Universal Robots PolyScope program: AdientTorsF_Eol1R.urp

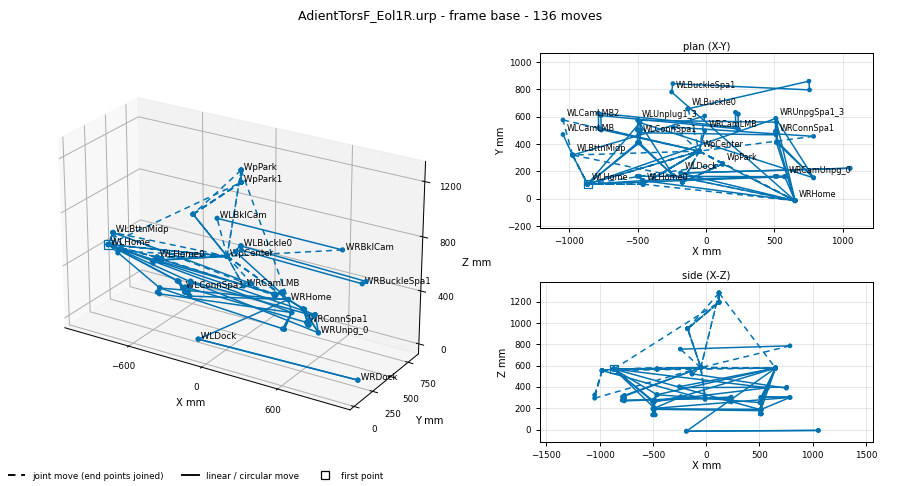
[picture p0: tool path of AdientTorsF_Eol1R.urp in frame base, 136 of 176 moves have a stored position in this frame; points joined in program order, loops and branches not executed]
Program AdientTorsF_Eol1R (installation=EOL_1R directory=/programs createdIn=3.5.1 lastSavedIn=5.26.0 robotSerialNumber=20265101874)
Calibrated DH parameters: a=[0.000042, -0.610949, -0.549442, -0.000024, -0.000005, 0]; d=[0.18065, -32.695743, 7.316343, 25.554022, 0.119806, 0.115349]; alpha=[1.570492, -0.001088, 0.006138, 1.570534, -1.57033, 0]; deltaTheta=[0, 0.058138, -0.334397, 0.276266, -0.000002, 0]
InitVariablesNode variables(variable(name=Abort, expression=False), variable(name=AdapterReady_L, expression=False), variable(name=AdapterReady_R, expression=False), variable(name=CMD_Heartbt_i1, expression=0), variable(name=CMD_Heartbt_i2, expression=0), variable(name=CMD_Program_i1, expression=0), variable(name=CMD_Program_i2, expression=0), variable(name=CMD_Reserve_i1, expression=0), variable(name=CMD_Reserve_i2, expression=0), variable(name=CMD_Timeout_i1, expression=0), variable(name=CMD_Timeout_i2, expression=0), variable(name=CamCorrectnOK, expression=0), variable(name=DEBUG, expression=False), variable(name=D_rel, expression=p[0,0,0,0,0,0]), variable(name=EvtBeep, expression=False), variable(name=EvtDock, expression=0), variable(name=Mute, expression=False), variable(name=P_ini, expression=get_actual_tcp_pose()), variable(name=Parking, expression=0), variable(name=ProgExe, expression=0), variable(name=STS_Heartbeat, expression=False), variable(name=STS_Progress, expression=0), variable(name=STS_Reservation, expression=0), variable(name=SetCameraProg, expression=0))
BeforeStart
  SuppressedNode
    DEBUG := True
  'SW version, to be used to track changes and keep sync of all stations'
  SW_Ver := 1.0
  Folder Scripts [hidden by the author, left out]
  Folder Avoid guidance screen [hidden by the author, left out]
  Call GripperOpen
  GoToHome := True
  Script: socket_open("127.0.0.1",30001)
Robot Program (runOnlyOnce=false)
  Folder Execute Program
    Folder Init
      Wait Condition expression=EvtDock≤0
      Folder Verify adapter ready
        If Di_Docked_L or AI_Gripper<(ivGripSensOpen+0.3)
          AdapterReady_L := False
        If Di_Docked_R or AI_Gripper<(ivGripSensOpen+0.3)
          AdapterReady_R := False
      Folder Go to home pos automatically
        If GoToHome and  not (AdapterReady_L or AdapterReady_R)
          Wait Sleep waitTime=1
          If InRange(P_Flange[0],-1,-0.2) and InRange(P_Flange[1],-0.5,0.5) and InRange(P_Flange[2],0.3,1)
            If AdapterDocked or DEBUG or (AI_Gripper<(ivGripSensOpen+0.3))
              MoveJ speed 120 deg/s, acceleration 500 deg/s^2 (useActiveTCP=false positionType=JointAngles optimoveEnabled=false optiMoveSpeed=0.3 optiMoveAcceleration=0.09) tcp=t0_Flange; feature=Base
                Waypoint WLHome: TCP in base x=-866.235 y=106.553 z=568.537 mm, rx=3.1416 ry=0 rz=0 rad; joints [-18.569, -73.864, 82.281, -98.358, -89.699, -108.526] deg; TCP offset x=0 y=0 z=0 mm, rx=0 ry=0 rz=3.1416 rad
            Else 
              Popup Error (haltProgram=false message=Adapter must be docked inputType=Text)
              Halt
          ElseIf AtCenterPos
            MoveJ speed 120 deg/s, acceleration 500 deg/s^2 (useActiveTCP=true positionType=JointAngles optimoveEnabled=false optiMoveSpeed=0.3 optiMoveAcceleration=0.09) feature=Base
              Waypoint WpCenter: TCP in base x=-50 y=348.529 z=581.932 mm, rx=0 ry=3.1416 rz=0 rad; joints [-111.545, -128.858, 124.717, -85.8, -89.657, -21.591] deg; TCP offset x=0 y=0 z=0 mm, rx=0 ry=0 rz=3.1416 rad
          ElseIf AtParkPos
            MoveJ speed 120 deg/s, acceleration 500 deg/s^2 (useActiveTCP=true positionType=JointAngles optimoveEnabled=false optiMoveSpeed=0.3 optiMoveAcceleration=0.09) feature=Base
              Waypoint WpPark: TCP in base x=121.203 y=255.21 z=1282.913 mm, rx=-1.7636 ry=-1.7554 rz=-0.7332 rad; joints [-180, -89.998, -0.001, 0.001, -45, 0] deg; TCP offset x=0 y=0 z=0 mm, rx=0 ry=0 rz=3.1416 rad
          ElseIf InRange(P_Flange[0],0.2,1.2) and InRange(P_Flange[1],-0.5,0.5) and InRange(P_Flange[2],0.3,1)
            If AdapterDocked or DEBUG or (AI_Gripper<(ivGripSensOpen+0.3))
              MoveJ speed 120 deg/s, acceleration 500 deg/s^2 (useActiveTCP=true positionType=JointAngles optimoveEnabled=false optiMoveSpeed=0.3 optiMoveAcceleration=0.09) feature=Base
                Waypoint WRHome: TCP in base x=651.404 y=-14.037 z=577.942 mm, rx=3.1416 ry=0 rz=0 rad; joints [-196.798, -95.185, 104.834, -99.59, -89.673, 73.253] deg
            Else 
              Popup Error (haltProgram=false message=Adapter must be docked inputType=Text)
              Halt
          Else 
            Popup Error (haltProgram=false message=Illegal position. Adjust arm to open space in front of the backrest, or [Move]->[Home] inputType=Text)
            Halt
        GoToHome := False
      If DEBUG
        'Popup window with program selection'
        ProgExe :=  (valueSource=Operator message=Program number? valueType=Integer)
      If ProgExe>0
        Folder Init
          Mute := False
          Wait Condition expression=not GoToHome
          If In(ProgExe,[11,12,14])
            AdapterReady_R := False
          ElseIf In(ProgExe,[51,52,54])
            AdapterReady_L := False
          Else 
            AdapterReady_L := False
            AdapterReady_R := False
    Folder Programs
      If InRange(ProgExe,1,99)
        Folder Undock
          If In(ProgExe,[11,51])
            Script: Report(1)
            Folder AtHome?
              Timer (action=Reset) variable(name=T_Timeout)
              Timer (action=Start) variable=T_Timeout
              Wait Condition expression=AtHomePos or T_Timeout>5
              If not AtHomePos
                Script: Report(90)
            If Progress_run() and  not AdapterDocked
              Script: Report(94)
            If Progress_run()
              Folder Undock
                MoveL speed 1000 mm/s, acceleration 3000 mm/s^2 (useActiveTCP=false optimoveEnabled=false optiMoveSpeed=0.3 optiMoveAcceleration=0.09) tcp=t2_Gripper; feature=Base
                  Call GripperOpenQuick
                  If False
                    Waypoint WLDock: TCP in base x=-185.159 y=188.226 z=-15.087 mm, rx=1.8903 ry=-1.8549 rz=-0.6082 rad; joints [-63.281, -90.699, 161.642, -179.168, -58.985, -58.884] deg; TCP offset x=0 y=260 z=74 mm, rx=0 ry=0 rz=3.1416 rad
                    Waypoint WRDock: TCP in base x=1053.302 y=223.512 z=-7.7 mm, rx=1.9028 ry=-1.8549 rz=-0.594 rad; joints [-177.46, -52.491, 84.331, -87.181, -88.23, 180.6] deg
                  If ProgExe<50
                    WpDock := WLDock
                    WpHome := WLHome
                  Else 
                    WpDock := WRDock
                    WpHome := WRHome
                  Wp := pose_trans(WpDock, p[0,0.175,-0.1,0,0,0])
                  Waypoint Variable (Variable): motionParameters(blendRadius=0.05); variable=Wp
                  Call GripperOpen
                  Wp := pose_trans(WpDock, p[0,0.075,0.01,0,0,0])
                  Waypoint Variable (Variable): motionParameters(blendRadius=0.01); variable=Wp
                  Wp := pose_trans(WpDock, p[0,0.055,0,0,0,0])
                  Waypoint Variable (Variable): motionParameters(blendRadius=0.01); variable=Wp
                  Waypoint Variable (Variable): variable=WpDock
                  Call GripperClose
                  Wp := pose_trans(WpDock, p[0,0.25,0,0,0,0])
                  Waypoint Variable (Variable): variable=Wp
                If ProgExe<50
                  AdapterReady_L := True
                Else 
                  AdapterReady_R := True
                Script: Report(50)
            Script: Report(50)
        Folder Connect
          If In(ProgExe,[12,14,52,54])
            Script: Report(1)
            If ProgExe<50 and AdapterReady_L
              Undock := False
            ElseIf ProgExe≥50 and AdapterReady_R
              Undock := False
            Else 
              Undock := True
              Folder AtHome? [hidden by the author, left out]
              If Progress_run() and  not AdapterDocked
                Script: Report(94)
            If Progress_run()
              Folder Undock
                If Undock
                  MoveL speed 1000 mm/s, acceleration 3000 mm/s^2 (useActiveTCP=false optimoveEnabled=false optiMoveSpeed=0.3 optiMoveAcceleration=0.09) tcp=t2_Gripper; feature=Base
                    Call GripperOpenQuick
                    If False
                      Waypoint WLDock: TCP in base x=-185.159 y=188.226 z=-15.087 mm, rx=1.8903 ry=-1.8549 rz=-0.6082 rad; joints [-63.281, -90.699, 161.642, -179.168, -58.985, -58.884] deg; TCP offset x=0 y=260 z=74 mm, rx=0 ry=0 rz=3.1416 rad
                      Waypoint WRDock: TCP in base x=1053.302 y=223.512 z=-7.7 mm, rx=1.9028 ry=-1.8549 rz=-0.594 rad; joints [-177.46, -52.491, 84.331, -87.181, -88.23, 180.6] deg
                    If ProgExe<50
                      WpDock := WLDock
                      WpHome := WLHome
                    Else 
                      WpDock := WRDock
                      WpHome := WRHome
                    Wp := pose_trans(WpDock, p[0,0.175,-0.1,0,0,0])
                    Waypoint Variable (Variable): motionParameters(blendRadius=0.05); variable=Wp
                    Call GripperOpen
                    Wp := pose_trans(WpDock, p[0,0.075,0.01,0,0,0])
                    Waypoint Variable (Variable): motionParameters(blendRadius=0.01); variable=Wp
                    Wp := pose_trans(WpDock, p[0,0.055,0,0,0,0])
                    Waypoint Variable (Variable): motionParameters(blendRadius=0.01); variable=Wp
                    Waypoint Variable (Variable): variable=WpDock
                    Call GripperClose
                    Wp := pose_trans(WpDock, p[0,0.25,0,0,0,0])
                    Waypoint Variable (Variable): variable=Wp
                AdapterReady_L := False
                AdapterReady_R := False
                Script: Report(2)
              CamCorrection := p[0,0,0,0,0,0]
              SuppressedNode
                Folder Camera
                  MoveL speed 250 mm/s, acceleration 1200 mm/s^2 (useActiveTCP=false optimoveEnabled=false optiMoveSpeed=0.3 optiMoveAcceleration=0.09) tcp=t0_Flange; feature=Base
                    If In(ProgExe,[12,13])
                      SetCameraProg := 12
                      Waypoint WLCamConSpa1: TCP in base x=-511.083 y=256.44 z=253.227 mm, rx=2.1948 ry=2.1949 rz=-0.0574 rad; joints [170.312, -93.988, -133.728, -42.837, 93.248, -9.279] deg; TCP offset x=0 y=0 z=0 mm, rx=0 ry=0 rz=0 rad
                    If In(ProgExe,[14])
                      SetCameraProg := ProgExe
                      Waypoint WLCamConSpa3: TCP in base x=-559.049 y=229.366 z=263.196 mm, rx=-2.2214 ry=-2.2215 rz=0 rad; joints [174.302, -95.829, -130.307, -43.928, 90.296, -5.276] deg
                    If In(ProgExe,[52,53])
                      SetCameraProg := 52
                      Waypoint WRCamConSpa1: TCP in base x=528.577 y=256.538 z=254.589 mm, rx=2.1946 ry=2.1948 rz=-0.0575 rad; joints [43.439, -94.974, -131.929, -45.242, 88.117, 223.892] deg
                    If In(ProgExe,[54])
                      SetCameraProg := ProgExe
                      Waypoint WRCamConSpa3: TCP in base x=480.455 y=221.374 z=266.967 mm, rx=-2.2214 ry=-2.2215 rz=-0.0001 rad; joints [43.801, -88.335, -137.68, -44.047, 90.305, 224.222] deg
                  Call CamAcquire
                  CamCorrection := p[CamData[0],CamData[1]*-0.5,CamData[1],0,0,0]
            SuppressedNode
              If Progress_run() and CamCorrectnOK≠ProgExe
                EvtDock := 1
                Wait Condition expression=EvtDock≟0
                Script: Report(91)
            Folder Connect
              If Progress_run()
                Set NoAction tcp=t2_Gripper
                MoveL speed 1000 mm/s, acceleration 3000 mm/s^2 (useActiveTCP=false optimoveEnabled=false optiMoveSpeed=0.3 optiMoveAcceleration=0.09) tcp=t2_Gripper; feature=Base
                  If False
                    'wp is set to position exactly 30mm below'
                    Waypoint WLConnSpa1: motionParameters(blendRadius=0.013); TCP in base x=-494.014 y=464.207 z=189.073 mm, rx=3.1414 ry=0 rz=0 rad; joints [-41.576, -90.764, 137.111, -136.317, -89.71, -131.321] deg; TCP offset x=0 y=260 z=74 mm, rx=0 ry=0 rz=3.1416 rad
                    Waypoint WLConnSpa3: TCP in base x=-485.347 y=483.182 z=190.434 mm, rx=-3.1063 ry=0 rz=0 rad; joints [-43.288, -89.958, 137.919, -139.316, -91.202, -133.036] deg; TCP offset x=0 y=260 z=74 mm, rx=0 ry=0 rz=3.1416 rad
                    Waypoint WRConnSpa1: TCP in base x=512.219 y=467.564 z=177.585 mm, rx=3.1416 ry=0.0001 rz=-0.0002 rad; joints [-176.409, -87.84, 135.834, -137.962, -89.727, 93.852] deg; TCP offset x=0 y=260 z=74 mm, rx=0 ry=0 rz=3.1416 rad
                    Waypoint WRConnSpa3: TCP in base x=517.873 y=489.304 z=184.649 mm, rx=3.1416 ry=0.0001 rz=-0.0002 rad; joints [-174.123, -87.241, 134.145, -136.871, -89.724, 96.132] deg; TCP offset x=0 y=260 z=74 mm, rx=0 ry=0 rz=3.1416 rad
                  If In(ProgExe,[12])
                    Wp := pose_trans(WLConnSpa1, CamCorrection)
                  If In(ProgExe,[14])
                    Wp := pose_add(WLConnSpa3, CamCorrection)
                  If In(ProgExe,[52])
                    Wp := pose_trans(WRConnSpa1, CamCorrection)
                  If In(ProgExe,[54])
                    Wp := pose_add(WRConnSpa3, CamCorrection)
                  Waypoint Variable (Variable): variable=Wp
                Force Frame feature=Joint_6_name; selection=[0, 0, 1, 0, 0, 0]; wrench=[0, 0, -30, 0, 0, 0]; limitsForce=[0.15, 0.15, 0.1, 1.047198, 1.047198, 1.047198]; limitsMotion=[0.1, 0.1, 0.1, 0.349066, 0.349066, 0.349066]
                  Wait Sleep waitTime=1
                Force Frame feature=Joint_6_name; selection=[1, 0, 1, 0, 0, 0]; wrench=[0, 0, -30, 0, 0, 0]; limitsForce=[0.15, 0.15, 0.05, 1.047198, 1.047198, 1.047198]; limitsMotion=[0.1, 0.1, 0.1, 0.349066, 0.349066, 0.349066]
                  Wait Sleep waitTime=0.5
                'position ok'
                If InRange(Wp[2]+0.03-P_act[2],-0.015,0.015)
                  'ok'
                Else 
                  EvtDock := 2
                  Wait Condition expression=EvtDock≤0
                  Script: Report(96)
              If Progress_run()
                Force Frame feature=Joint_6_name; selection=[0, 1, 0, 0, 0, 0]; wrench=[0, -60, -10, 0, 0, 0]; limitsForce=[0.15, 0.05, 0.01, 1.047198, 1.047198, 1.047198]; limitsMotion=[0.1, 0.1, 0.1, 0.349066, 0.349066, 0.349066]
                  Wait Sleep waitTime=1
                MoveL speed 1000 mm/s, acceleration 3000 mm/s^2 (useActiveTCP=true optimoveEnabled=false optiMoveSpeed=0.3 optiMoveAcceleration=0.09) feature=Base
                  Wp := pose_trans(P_act, p[0,0.005,0,0,0,0])
                  Waypoint Variable (Variable): variable=Wp
                Call GripperOpen
                Force Frame feature=Joint_6_name; selection=[0, 1, 0, 0, 0, 0]; wrench=[0, -60, -10, 0, 0, 0]; limitsForce=[0.15, 0.1, 0.01, 1.047198, 1.047198, 1.047198]; limitsMotion=[0.1, 0.1, 0.1, 0.349066, 0.349066, 0.349066]
                  Wait Sleep waitTime=1
                  Script: Report(5)
                  MoveL speed 500 mm/s, acceleration 2000 mm/s^2 (useActiveTCP=true optimoveEnabled=false optiMoveSpeed=0.3 optiMoveAcceleration=0.09) feature=Base
                    Wp0 := get_actual_tcp_pose()
                    Wp := pose_trans(Wp0, p[0,0,0,0,0,0.07])
                    Waypoint Variable (Variable): variable=Wp
                    Wp := pose_trans(Wp0, p[0,0,0,0,0,-0.07])
                    Waypoint Variable (Variable): variable=Wp
                    Waypoint Variable (Variable): variable=Wp0
                    Wp := pose_trans(Wp0, p[0,0,0.01,0,0,0])
                    Waypoint Variable (Variable): variable=Wp
                    Waypoint Variable (Variable): variable=Wp0
                MoveL speed 1000 mm/s, acceleration 3000 mm/s^2 (useActiveTCP=true optimoveEnabled=false optiMoveSpeed=0.3 optiMoveAcceleration=0.09) feature=Base
                  Wp0 := get_actual_tcp_pose()
                  Wp := pose_trans(Wp0, p[0,0.015,0,0,0,0])
                  Waypoint Variable (Variable): variable=Wp
                Force Frame feature=Joint_6_name; selection=[0, 1, 0, 0, 0, 0]; wrench=[0, -60, 0, 0, 0, 0]; limitsForce=[0.15, 0.5, 0.15, 1.047198, 1.047198, 1.047198]; limitsMotion=[0.1, 0.1, 0.1, 0.349066, 0.349066, 0.349066]
                  Wait Sleep waitTime=0.5
                Script: Report(6)
                Timer (action=Reset) variable=T_Timeout
                Timer (action=Start) variable=T_Timeout
                Folder Test switch pin, retreat on fail
                  Wait Condition expression=Flags[0] or T_Timeout>10 or DEBUG
                  If not Flags[0] and  not DEBUG
                    EvtDock := 2
                    Wait Condition expression=EvtDock≤0
                    Script: Report(95)
            If Progress_run()
              MoveL speed 1000 mm/s, acceleration 3000 mm/s^2 (useActiveTCP=false optimoveEnabled=false optiMoveSpeed=0.3 optiMoveAcceleration=0.09) tcp=t0_Flange; feature=Base
                Set NoAction tcp=t0_Flange
                P_act := get_actual_tcp_pose()
                Wp := pose_trans(P_act, p[0,0.1,0,0,0,0])
                Waypoint Variable (Variable): motionParameters(blendRadius=0.05); variable=Wp
                Wp := pose_trans(Wp, p[0,0.1,-0.1,0,0,0])
                Waypoint Variable (Variable): motionParameters(blendRadius=0.05); variable=Wp
                Waypoint Variable (Variable): variable=WpHome
              Script: Report(50)
        Folder Buckle
          If In(ProgExe,[15,16,55,56])
            Script: Report(1)
            Folder AtHome?
              Timer (action=Reset) variable=T_Timeout
              Timer (action=Start) variable=T_Timeout
              Wait Condition expression=AtHomePos or (In(ProgExe,[15,16]) and AtCenterPos) or T_Timeout>5
              If AtHomePos or (In(ProgExe,[15,16]) and AtCenterPos)
                'nop'
              Else 
                Script: Report(90)
            If Progress_run() and  not ((Di_SBR_L_X_Wp and ProgExe<50)  or (Di_SBR_R_X_Wp and ProgExe>50))
              Script: Report(92)
            If Progress_run()
              Call GripperCloseQuick
              Folder Camera
                SetCameraProg := ProgExe
                MoveL speed 1000 mm/s, acceleration 3000 mm/s^2 (useActiveTCP=false optimoveEnabled=false optiMoveSpeed=0.3 optiMoveAcceleration=0.09) tcp=t0_Flange; feature=Base
                  If ProgExe<50
                    MoveJ speed 120 deg/s, acceleration 500 deg/s^2 (useActiveTCP=false positionType=JointAngles optimoveEnabled=false optiMoveSpeed=0.3 optiMoveAcceleration=0.09) tcp=t0_Flange; feature=Base
                      If AtLHomePos
                        Waypoint WLHome0: motionParameters(blendRadius=0.05); TCP in base x=-460.734 y=106.553 z=568.537 mm, rx=-2.2214 ry=2.2214 rz=0 rad; joints [-34.699, -114.011, 119.5, -95.429, -89.656, -34.68] deg; TCP offset x=0 y=0 z=0 mm, rx=0 ry=0 rz=3.1416 rad
                        Waypoint WpCenter: motionParameters(blendRadius=0.1); TCP in base x=-50 y=348.529 z=581.932 mm, rx=0 ry=3.1416 rz=0 rad; joints [-111.545, -128.858, 124.717, -85.8, -89.657, -21.591] deg; TCP offset x=0 y=0 z=0 mm, rx=0 ry=0 rz=3.1416 rad
                      Waypoint WLBklCam: TCP in base x=-241.801 y=524.603 z=755.343 mm, rx=0.5219 ry=-1.5373 rz=-0.5328 rad; joints [-95.3, -98.197, 89.288, -6.269, -4.596, -113.342] deg; TCP offset x=0 y=0 z=0 mm, rx=0 ry=0 rz=3.1416 rad
                  Else 
                    Waypoint WRBklCam: TCP in base x=786.942 y=456.735 z=786.447 mm, rx=-1.8153 ry=0.6794 rz=-1.6469 rad; joints [-158.937, -69.521, 77.508, -184.213, -106.091, 137.333] deg
                Call GripperClose
                Call CamAcquire
                Call CamCalculateCorectnPlane
              If CamCorrectnOK≟ProgExe and InRange(CamCorrection[1],-0.05,0.052) and InRange(CamCorrection[2],-0.03,0.03)
                'empty'
              Else 
                CamCorrectnOK := 0
                MoveJ speed 120 deg/s, acceleration 500 deg/s^2 (useActiveTCP=false positionType=JointAngles optimoveEnabled=false optiMoveSpeed=0.3 optiMoveAcceleration=0.09) tcp=t0_Flange; feature=Base
                  If ProgExe<50
                    MoveJ speed 180 deg/s, acceleration 1000 deg/s^2 (useActiveTCP=false positionType=JointAngles optimoveEnabled=false optiMoveSpeed=0.3 optiMoveAcceleration=0.09) tcp=t0_Flange; feature=Base
                      Waypoint WpCenter: TCP in base x=-50 y=348.529 z=581.932 mm, rx=0 ry=3.1416 rz=0 rad; joints [-111.545, -128.858, 124.717, -85.8, -89.657, -21.591] deg; TCP offset x=0 y=0 z=0 mm, rx=0 ry=0 rz=3.1416 rad
                      STS_Reservation := 0
                  Else 
                    Waypoint WRHome: TCP in base x=651.404 y=-14.037 z=577.942 mm, rx=3.1416 ry=0 rz=0 rad; joints [-196.798, -95.185, 104.834, -99.59, -89.673, 73.253] deg; TCP offset x=0 y=0 z=0 mm, rx=0 ry=0 rz=3.1416 rad
                Script: Report(91)
              If CamCorrectnOK≟ProgExe
                Folder Insert
                  MoveL speed 1000 mm/s, acceleration 3000 mm/s^2 (useActiveTCP=false optimoveEnabled=false optiMoveSpeed=0.3 optiMoveAcceleration=0.09) tcp=t3_Blade; feature=Base
                    If False
                      'must be set with blade ca one half into buckle slot'
                      Waypoint WLBuckleSpa1: TCP in base x=-251.61 y=780.85 z=402.619 mm, rx=-2.5257 ry=-0.026 rz=-0.03 rad; joints [-95.327, -89.75, 121.006, -156.476, -87.65, -185.489] deg; TCP offset x=134 y=56 z=118 mm, rx=0 ry=0 rz=-3.1416 rad
                      Waypoint WLBuckleSpa3: TCP in base x=-242.615 y=842.237 z=394.859 mm, rx=-2.618 ry=0 rz=0 rad; joints [-95.692, -84.24, 113.52, -149.146, -86.956, -184.638] deg
                      Waypoint WRBuckleSpa1: TCP in base x=756.879 y=796.528 z=397.405 mm, rx=-2.6367 ry=-0.0043 rz=-0.0316 rad; joints [-153.635, -49.484, 59.406, -114.921, -64.657, 119.621] deg
                      Waypoint WRBuckleSpa3: TCP in base x=752.503 y=860.244 z=388.844 mm, rx=-2.618 ry=0.0001 rz=0 rad; joints [-150.822, -45.037, 53.33, -114.028, -63.84, 122.901] deg
                    If ProgExe≟15
                      Wp := WLBuckleSpa1
                      Waypoint WLBuckle0: motionParameters(blendRadius=0.1); TCP in base x=-131.782 y=658.01 z=522.985 mm, rx=2.2703 ry=-2.1715 rz=0 rad; joints [-89.222, -105.834, 107.036, -91.142, -89.67, -91.771] deg; TCP offset x=134 y=56 z=118 mm, rx=0 ry=0 rz=-3.1416 rad
                    If ProgExe≟16
                      Wp := WLBuckleSpa3
                      Waypoint WLBuckle0: motionParameters(blendRadius=0.1); TCP in base x=-131.782 y=658.01 z=522.985 mm, rx=2.2703 ry=-2.1715 rz=0 rad; joints [-89.222, -105.834, 107.036, -91.142, -89.67, -91.771] deg
                    If ProgExe≟55
                      Wp := WRBuckleSpa1
                    If ProgExe≟56
                      Wp := WRBuckleSpa3
                    Wp0 := pose_trans(Wp,p[0,0,-0.02,0,0,0])
                    Wp0 := pose_add(Wp0,Base_w_correctn)
                    Waypoint Variable (Variable): variable=Wp0
                  Script: Report(5)
                  Timer (action=Reset) variable=T_Timeout
                  Timer (action=Start) variable=T_Timeout
                  Wait Condition expression=Flags[8] or Abort or DEBUG or T_Timeout>25
                  If Flags[8] or DEBUG
                    Script: Report(6)
                    Set NoAction tcp=t3_Blade
                    Force Frame feature=Joint_6_name; selection=[0, 0, 1, 0, 0, 0]; wrench=[0, 0, 15, 0, 0, 0]; limitsForce=[0.15, 0.15, 0.15, 1.047198, 1.047198, 1.047198]; limitsMotion=[0.1, 0.1, 0.1, 0.349066, 0.349066, 0.349066]
                      Wait Sleep waitTime=1
                    If not Flags[9] and  not Abort
                      MoveL speed 50 mm/s, acceleration 500 mm/s^2 (useActiveTCP=false optimoveEnabled=false optiMoveSpeed=0.3 optiMoveAcceleration=0.09) tcp=t3_Blade; feature=Base
                        Waypoint Variable (Variable): variable=Wp
                      Force Frame feature=Joint_6_name; selection=[1, 1, 1, 0, 0, 0]; wrench=[0, 0, 50, 0, 0, 0]; limitsForce=[0.15, 0.15, 0.25, 1.047198, 1.047198, 1.047198]; limitsMotion=[0.1, 0.1, 0.1, 0.349066, 0.349066, 0.349066]
                        Wait Sleep waitTime=1.5
                    If not Flags[9] and  not Abort
                      MoveL speed 50 mm/s, acceleration 500 mm/s^2 (useActiveTCP=false optimoveEnabled=false optiMoveSpeed=0.3 optiMoveAcceleration=0.09) tcp=t3_Blade; feature=Base
                        Waypoint Variable (Variable): variable=Wp
                      Force Frame feature=Joint_6_name; selection=[1, 1, 1, 0, 0, 0]; wrench=[0, 0, 50, 0, 0, 0]; limitsForce=[0.15, 0.15, 0.25, 1.047198, 1.047198, 1.047198]; limitsMotion=[0.1, 0.1, 0.1, 0.349066, 0.349066, 0.349066]
                        Wait Sleep waitTime=1.5
                    If not Flags[9] and  not Abort
                      MoveL speed 50 mm/s, acceleration 500 mm/s^2 (useActiveTCP=false optimoveEnabled=false optiMoveSpeed=0.3 optiMoveAcceleration=0.09) tcp=t3_Blade; feature=Base
                        Waypoint Variable (Variable): variable=Wp
                      Force Frame feature=Joint_6_name; selection=[1, 1, 1, 0, 0, 0]; wrench=[0, 0, 50, 0, 0, 0]; limitsForce=[0.15, 0.15, 0.25, 1.047198, 1.047198, 1.047198]; limitsMotion=[0.1, 0.1, 0.1, 0.349066, 0.349066, 0.349066]
                        Wait Sleep waitTime=1.5
                  MoveL speed 1000 mm/s, acceleration 3000 mm/s^2 (useActiveTCP=false optimoveEnabled=false optiMoveSpeed=0.3 optiMoveAcceleration=0.09) tcp=t3_Blade; feature=Base
                    Waypoint Variable (Variable): variable=Wp
                    MoveDirectionNode (selectedDirection=ZMinus) feature=Joint_6_name
                      Until DISTANCE (allowActions=false deceleration=3 distanceNodeType=STOP) Distance=0.02; motionParameters(blendRadius=0)
                    If In(ProgExe,[15,16])
                      MoveJ speed 180 deg/s, acceleration 1000 deg/s^2 (useActiveTCP=false positionType=JointAngles optimoveEnabled=false optiMoveSpeed=0.3 optiMoveAcceleration=0.09) tcp=t0_Flange; feature=Base
                        Waypoint WLBuckle0: motionParameters(blendRadius=0.1); TCP in base x=-131.782 y=658.01 z=522.985 mm, rx=2.2703 ry=-2.1715 rz=0 rad; joints [-89.222, -105.834, 107.036, -91.142, -89.67, -91.771] deg; TCP offset x=134 y=56 z=118 mm, rx=0 ry=0 rz=-3.1416 rad
                        Waypoint WpCenter: TCP in base x=-50 y=348.529 z=581.932 mm, rx=0 ry=3.1416 rz=0 rad; joints [-111.545, -128.858, 124.717, -85.8, -89.657, -21.591] deg; TCP offset x=0 y=0 z=0 mm, rx=0 ry=0 rz=3.1416 rad
                        STS_Reservation := 0
                    If In(ProgExe,[55,56])
                      MoveJ speed 120 deg/s, acceleration 500 deg/s^2 (useActiveTCP=false positionType=JointAngles optimoveEnabled=false optiMoveSpeed=0.3 optiMoveAcceleration=0.09) tcp=t0_Flange; feature=Base
                        Waypoint WRHome: TCP in base x=651.404 y=-14.037 z=577.942 mm, rx=3.1416 ry=0 rz=0 rad; joints [-196.798, -95.185, 104.834, -99.59, -89.673, 73.253] deg; TCP offset x=0 y=0 z=0 mm, rx=0 ry=0 rz=3.1416 rad
                  If Progress_check()≥6
                    Script: Report(50)
                  Else 
                    Script: Report(95)
        Folder Disconnect
          If In(ProgExe,[21,22,23,61,62,63])
            Script: Report(1)
            Folder AtHome? [hidden by the author, left out]
            If Progress_run()
              If In(ProgExe,[21,22])
                SetCameraProg := 21
                MoveL speed 1000 mm/s, acceleration 3000 mm/s^2 (useActiveTCP=false optimoveEnabled=false optiMoveSpeed=0.3 optiMoveAcceleration=0.09) tcp=t0_Flange; feature=Base
                  Waypoint WLCamUnpg_0: motionParameters(blendRadius=0.05); TCP in base x=-461.191 y=133.026 z=327.436 mm, rx=2.2214 ry=-2.2214 rz=0 rad; joints [-37.473, -102.86, 138.571, -125.652, -89.683, -37.272] deg
                  Waypoint WLCamUnplgSpa1: TCP in base x=-503.393 y=164.68 z=272.56 mm, rx=2.163 ry=-2.163 rz=0.1228 rad; joints [-38.596, -92.511, 136.321, -129.705, -84.623, -38.554] deg
              If In(ProgExe,[23])
                SetCameraProg := ProgExe
                MoveL speed 1000 mm/s, acceleration 3000 mm/s^2 (useActiveTCP=false optimoveEnabled=false optiMoveSpeed=0.3 optiMoveAcceleration=0.09) tcp=t0_Flange; feature=Base
                  Waypoint WLCamUnpg_0: motionParameters(blendRadius=0.05); TCP in base x=-461.191 y=133.026 z=327.436 mm, rx=2.2214 ry=-2.2214 rz=0 rad; joints [-37.473, -102.86, 138.571, -125.652, -89.683, -37.272] deg
                  Waypoint WLCamUnpgSpa3: TCP in base x=-486.088 y=164.68 z=264.125 mm, rx=2.163 ry=-2.163 rz=0.1228 rad; joints [-39.861, -93.42, 138.312, -130.675, -84.715, -39.815] deg
              If In(ProgExe,[61,62])
                SetCameraProg := 61
                MoveL speed 1000 mm/s, acceleration 3000 mm/s^2 (useActiveTCP=false optimoveEnabled=false optiMoveSpeed=0.3 optiMoveAcceleration=0.09) tcp=t0_Flange; feature=Base
                  Waypoint WRCamUnpg_0: motionParameters(blendRadius=0.05); TCP in base x=575.167 y=161.724 z=392.695 mm, rx=-2.2214 ry=2.2214 rz=0 rad; joints [-181.33, -94.222, 123.788, -119.507, -89.682, 178.838] deg; TCP offset x=0 y=0 z=0 mm, rx=0 ry=0 rz=3.1416 rad
                  Waypoint WRCamUnplgSpa1: TCP in base x=505.675 y=163.851 z=252.755 mm, rx=2.163 ry=-2.163 rz=0.1228 rad; joints [-179.803, -89.572, 137.529, -137.844, -96.23, 180.476] deg; TCP offset x=0 y=0 z=0 mm, rx=0 ry=0 rz=3.1416 rad
              If In(ProgExe,[63])
                SetCameraProg := ProgExe
                MoveL speed 1000 mm/s, acceleration 3000 mm/s^2 (useActiveTCP=false optimoveEnabled=false optiMoveSpeed=0.3 optiMoveAcceleration=0.09) tcp=t0_Flange; feature=Base
                  Waypoint WRCamUnpg_0: motionParameters(blendRadius=0.05); TCP in base x=575.167 y=161.724 z=392.695 mm, rx=-2.2214 ry=2.2214 rz=0 rad; joints [-181.33, -94.222, 123.788, -119.507, -89.682, 178.838] deg; TCP offset x=0 y=0 z=0 mm, rx=0 ry=0 rz=3.1416 rad
                  Waypoint WRCamUnpgSpa3: TCP in base x=519.232 y=163.85 z=252.755 mm, rx=2.163 ry=-2.163 rz=0.1228 rad; joints [-179.81, -88.33, 136.25, -137.809, -96.231, 180.469] deg; TCP offset x=0 y=0 z=0 mm, rx=0 ry=0 rz=3.1416 rad
              Call CamAcquire
              Call CamCalculateCorectnPlane
            If Progress_run() and CamCorrectnOK≠ProgExe
              MoveL speed 1000 mm/s, acceleration 3000 mm/s^2 (useActiveTCP=false optimoveEnabled=false optiMoveSpeed=0.3 optiMoveAcceleration=0.09) tcp=t0_Flange; feature=Base
                If ProgExe<50
                  Waypoint WLCamUnpg_0: motionParameters(blendRadius=0.05); TCP in base x=-461.191 y=133.026 z=327.436 mm, rx=2.2214 ry=-2.2214 rz=0 rad; joints [-37.473, -102.86, 138.571, -125.652, -89.683, -37.272] deg
                  Waypoint WLHome: TCP in base x=-866.235 y=106.553 z=568.537 mm, rx=3.1416 ry=0 rz=0 rad; joints [-18.569, -73.864, 82.281, -98.358, -89.699, -108.526] deg
                Else 
                  Waypoint WRCamUnpg_0: motionParameters(blendRadius=0.05); TCP in base x=575.167 y=161.724 z=392.695 mm, rx=-2.2214 ry=2.2214 rz=0 rad; joints [-181.33, -94.222, 123.788, -119.507, -89.682, 178.838] deg; TCP offset x=0 y=0 z=0 mm, rx=0 ry=0 rz=3.1416 rad
                  Waypoint WRHome: TCP in base x=651.404 y=-14.037 z=577.942 mm, rx=3.1416 ry=0 rz=0 rad; joints [-196.798, -95.185, 104.834, -99.59, -89.673, 73.253] deg; TCP offset x=0 y=0 z=0 mm, rx=0 ry=0 rz=3.1416 rad
              Script: Report(91)
            If Progress_run()
              Call GripperOpenQuick
              Folder Disconnect
                If In(ProgExe,[21,22])
                  MoveL speed 1000 mm/s, acceleration 3000 mm/s^2 (useActiveTCP=false optimoveEnabled=false optiMoveSpeed=0.3 optiMoveAcceleration=0.09) tcp=t2_Gripper; feature=Base_w_correctn
                    Waypoint WLUnlplug_0: motionParameters(blendRadius=0.05); TCP in base x=-238.065 y=168.589 z=307.202 mm, rx=-2.2215 ry=2.2215 rz=0 rad; joints [-38.137, -101.279, 130.996, -119.658, -89.675, -37.97] deg; TCP offset x=0 y=260 z=74 mm, rx=0 ry=0 rz=3.1416 rad
                    Call GripperOpen
                    Waypoint WLUnplug1_1: motionParameters(blendRadius=0.05); TCP in base x=-500.466 y=409.772 z=262.286 mm, rx=3.1416 ry=0 rz=0 rad; joints [-36.238, -98.57, 134.242, -125.613, -89.687, -126.035] deg; TCP offset x=0 y=260 z=74 mm, rx=0 ry=0 rz=3.1416 rad
                    Waypoint WLUnplug1_2: motionParameters(blendRadius=0.05); TCP in base x=-500.464 y=502.943 z=138.784 mm, rx=2.6168 ry=0 rz=0 rad; joints [-52.954, -89.068, 121.74, -97.822, -72.083, -146.82] deg
                    Waypoint WLUnplug1_3: TCP in base x=-498.469 y=574.234 z=195.355 mm, rx=3.0223 ry=0 rz=0 rad; joints [-51.068, -88.164, 128.017, -124.513, -85.394, -141.077] deg
                If In(ProgExe,[23])
                  MoveL speed 1000 mm/s, acceleration 3000 mm/s^2 (useActiveTCP=false optimoveEnabled=false optiMoveSpeed=0.3 optiMoveAcceleration=0.09) tcp=t2_Gripper; feature=Base_w_correctn
                    Waypoint WLUnlplug_0: motionParameters(blendRadius=0.05); TCP in base x=-238.065 y=168.589 z=307.202 mm, rx=-2.2215 ry=2.2215 rz=0 rad; joints [-38.137, -101.279, 130.996, -119.658, -89.675, -37.97] deg; TCP offset x=0 y=260 z=74 mm, rx=0 ry=0 rz=3.1416 rad
                    Call GripperOpen
                    Waypoint WLUnplg3_1: motionParameters(blendRadius=0.05); TCP in base x=-487.566 y=409.773 z=262.286 mm, rx=3.1416 ry=0 rz=0 rad; joints [-37.146, -99.98, 135.351, -125.313, -89.685, -126.946] deg; TCP offset x=0 y=260 z=74 mm, rx=0 ry=0 rz=3.1416 rad
                    Waypoint WLUnplg3_2: motionParameters(blendRadius=0.005); TCP in base x=-479.036 y=502.944 z=138.784 mm, rx=2.6168 ry=0 rz=0 rad; joints [-54.611, -90.718, 123.3, -97.296, -72.776, -148.397] deg
                    Waypoint WLUnplg3_3: TCP in base x=-483.481 y=557.037 z=199.597 mm, rx=3.0989 ry=0.009 rz=0.0106 rad; joints [-50.109, -89.474, 132.186, -130.561, -88.44, -140.24] deg
                If In(ProgExe,[61,62])
                  MoveL speed 1000 mm/s, acceleration 3000 mm/s^2 (useActiveTCP=false optimoveEnabled=false optiMoveSpeed=0.3 optiMoveAcceleration=0.09) tcp=t2_Gripper; feature=Base_w_correctn
                    Waypoint WRUnpg_0: motionParameters(blendRadius=0.05); TCP in base x=786.992 y=153.256 z=301.741 mm, rx=2.2214 ry=-2.2214 rz=0 rad; joints [-182.381, -98.367, 129.337, -120.911, -89.68, 177.795] deg
                    Call GripperOpen
                    Waypoint WRUnpgSpa1_1: motionParameters(blendRadius=0.05); TCP in base x=526.991 y=413.255 z=301.742 mm, rx=3.1416 ry=0 rz=0 rad; joints [-182.381, -98.367, 129.337, -120.911, -89.679, 87.795] deg; TCP offset x=0 y=260 z=74 mm, rx=0 ry=0 rz=3.1416 rad
                    Waypoint WRUnpgSpa1_2: motionParameters(blendRadius=0.05); TCP in base x=508.368 y=493.367 z=148.04 mm, rx=2.6127 ry=0 rz=0.0001 rad; joints [-160.596, -88.642, 123.424, -113.695, -118.08, 112.354] deg; TCP offset x=0 y=260 z=74 mm, rx=0 ry=0 rz=3.1416 rad
                    Waypoint WRUnpgSpa1_3: motionParameters(blendRadius=0); TCP in base x=510.847 y=587.448 z=186.724 mm, rx=3.0661 ry=0 rz=0.0001 rad; joints [-162.699, -84.876, 128.14, -131.932, -93.839, 107.582] deg
                If In(ProgExe,[63])
                  MoveL speed 1000 mm/s, acceleration 3000 mm/s^2 (useActiveTCP=false optimoveEnabled=false optiMoveSpeed=0.3 optiMoveAcceleration=0.09) tcp=t2_Gripper; feature=Base_w_correctn
                    Waypoint WRUnpg_0: motionParameters(blendRadius=0.05); TCP in base x=786.992 y=153.256 z=301.741 mm, rx=2.2214 ry=-2.2214 rz=0 rad; joints [-182.381, -98.367, 129.337, -120.911, -89.68, 177.795] deg
                    Call GripperOpen
                    Waypoint WRUnpg3_1: motionParameters(blendRadius=0.05); TCP in base x=513.973 y=413.256 z=301.741 mm, rx=3.1414 ry=0 rz=0 rad; joints [-182.44, -99.749, 130.447, -120.639, -89.678, 87.733] deg
                    Waypoint WRUnpg3_2: motionParameters(blendRadius=0.05); TCP in base x=517.647 y=493.368 z=148.039 mm, rx=2.618 ry=0 rz=0 rad; joints [-161.032, -87.955, 122.871, -114.143, -117.89, 111.838] deg; TCP offset x=0 y=260 z=74 mm, rx=0 ry=0 rz=3.1416 rad
                    Waypoint WRUnpg3_3: TCP in base x=515.624 y=560.572 z=190.167 mm, rx=3.1077 ry=0.0556 rz=0.0009 rad; joints [-166.386, -84.764, 129.261, -134.079, -91.592, 101.815] deg; TCP offset x=0 y=260 z=74 mm, rx=0 ry=0 rz=3.1416 rad
                Script: Report(20)
                Wait Condition expression=Flags[7] or DEBUG
              EvtDock := 2
              Wait Condition expression=EvtDock≤0
              If EvtDock<0
                If In(ProgExe,[21,22])
                  MoveL speed 1000 mm/s, acceleration 3000 mm/s^2 (useActiveTCP=false optimoveEnabled=false optiMoveSpeed=0.3 optiMoveAcceleration=0.09) tcp=t2_Gripper; feature=Base_w_correctn
                    Waypoint WLUnplug1_3: TCP in base x=-498.469 y=574.234 z=195.355 mm, rx=3.0223 ry=0 rz=0 rad; joints [-51.068, -88.164, 128.017, -124.513, -85.394, -141.077] deg
                    Waypoint WLUnplug1_2: motionParameters(blendRadius=0); TCP in base x=-500.464 y=502.943 z=138.784 mm, rx=2.6168 ry=0 rz=0 rad; joints [-52.954, -89.068, 121.74, -97.822, -72.083, -146.82] deg
                    Waypoint WLUnplug1_1: TCP in base x=-500.466 y=409.772 z=262.286 mm, rx=3.1416 ry=0 rz=0 rad; joints [-36.238, -98.57, 134.242, -125.613, -89.687, -126.035] deg
                  MoveL speed 1000 mm/s, acceleration 3000 mm/s^2 (useActiveTCP=false optimoveEnabled=false optiMoveSpeed=0.3 optiMoveAcceleration=0.09) tcp=t0_Flange; feature=Base
                    Waypoint WLHome: TCP in base x=-866.235 y=106.553 z=568.537 mm, rx=3.1416 ry=0 rz=0 rad; joints [-18.569, -73.864, 82.281, -98.358, -89.699, -108.526] deg; TCP offset x=0 y=0 z=0 mm, rx=0 ry=0 rz=3.1416 rad
                If In(ProgExe,[23])
                  MoveL speed 1000 mm/s, acceleration 3000 mm/s^2 (useActiveTCP=false optimoveEnabled=false optiMoveSpeed=0.3 optiMoveAcceleration=0.09) tcp=t2_Gripper; feature=Base_w_correctn
                    Waypoint WLUnplg3_3: TCP in base x=-483.481 y=557.037 z=199.597 mm, rx=3.0989 ry=0.009 rz=0.0106 rad; joints [-50.109, -89.474, 132.186, -130.561, -88.44, -140.24] deg; TCP offset x=0 y=260 z=74 mm, rx=0 ry=0 rz=3.1416 rad
                    Waypoint WLUnplg3_2: TCP in base x=-479.036 y=502.944 z=138.784 mm, rx=2.6168 ry=0 rz=0 rad; joints [-54.611, -90.718, 123.3, -97.296, -72.776, -148.397] deg
                    Waypoint WLUnplg3_1: TCP in base x=-487.566 y=409.773 z=262.286 mm, rx=3.1416 ry=0 rz=0 rad; joints [-37.146, -99.98, 135.351, -125.313, -89.685, -126.946] deg
                  MoveL speed 1000 mm/s, acceleration 3000 mm/s^2 (useActiveTCP=false optimoveEnabled=false optiMoveSpeed=0.3 optiMoveAcceleration=0.09) tcp=t0_Flange; feature=Base
                    Waypoint WLHome: TCP in base x=-866.235 y=106.553 z=568.537 mm, rx=3.1416 ry=0 rz=0 rad; joints [-18.569, -73.864, 82.281, -98.358, -89.699, -108.526] deg; TCP offset x=0 y=0 z=0 mm, rx=0 ry=0 rz=3.1416 rad
                If In(ProgExe,[61,62])
                  MoveL speed 1000 mm/s, acceleration 3000 mm/s^2 (useActiveTCP=false optimoveEnabled=false optiMoveSpeed=0.3 optiMoveAcceleration=0.09) tcp=t2_Gripper; feature=Base_w_correctn
                    Waypoint WRUnpgSpa1_3: motionParameters(blendRadius=0); TCP in base x=510.847 y=587.448 z=186.724 mm, rx=3.0661 ry=0 rz=0.0001 rad; joints [-162.699, -84.876, 128.14, -131.932, -93.839, 107.582] deg; TCP offset x=0 y=260 z=74 mm, rx=0 ry=0 rz=3.1416 rad
                    Waypoint WRUnpgSpa1_2: motionParameters(blendRadius=0.03); TCP in base x=508.368 y=493.367 z=148.04 mm, rx=2.6127 ry=0 rz=0.0001 rad; joints [-160.596, -88.642, 123.424, -113.695, -118.08, 112.354] deg
                    Waypoint WRUnpgSpa1_1: TCP in base x=526.991 y=413.255 z=301.742 mm, rx=3.1416 ry=0 rz=0 rad; joints [-182.381, -98.367, 129.337, -120.911, -89.679, 87.795] deg; TCP offset x=0 y=260 z=74 mm, rx=0 ry=0 rz=3.1416 rad
                  MoveL speed 1000 mm/s, acceleration 3000 mm/s^2 (useActiveTCP=false optimoveEnabled=false optiMoveSpeed=0.3 optiMoveAcceleration=0.09) tcp=t0_Flange; feature=Base
                    Waypoint WRHome: TCP in base x=651.404 y=-14.037 z=577.942 mm, rx=3.1416 ry=0 rz=0 rad; joints [-196.798, -95.185, 104.834, -99.59, -89.673, 73.253] deg; TCP offset x=0 y=0 z=0 mm, rx=0 ry=0 rz=3.1416 rad
                If In(ProgExe,[63])
                  MoveL speed 1000 mm/s, acceleration 3000 mm/s^2 (useActiveTCP=false optimoveEnabled=false optiMoveSpeed=0.3 optiMoveAcceleration=0.09) tcp=t2_Gripper; feature=Base_w_correctn
                    Waypoint WRUnpg3_3: TCP in base x=515.624 y=560.572 z=190.167 mm, rx=3.1077 ry=0.0556 rz=0.0009 rad; joints [-166.386, -84.764, 129.261, -134.079, -91.592, 101.815] deg; TCP offset x=0 y=260 z=74 mm, rx=0 ry=0 rz=3.1416 rad
                    Waypoint WRUnpg3_2: TCP in base x=517.647 y=493.368 z=148.039 mm, rx=2.618 ry=0 rz=0 rad; joints [-161.032, -87.955, 122.871, -114.143, -117.89, 111.838] deg; TCP offset x=0 y=260 z=74 mm, rx=0 ry=0 rz=3.1416 rad
                    Waypoint WRUnpg3_1: TCP in base x=513.973 y=413.256 z=301.741 mm, rx=3.1414 ry=0 rz=0 rad; joints [-182.44, -99.749, 130.447, -120.639, -89.678, 87.733] deg; TCP offset x=0 y=260 z=74 mm, rx=0 ry=0 rz=3.1416 rad
                  MoveL speed 1000 mm/s, acceleration 3000 mm/s^2 (useActiveTCP=false optimoveEnabled=false optiMoveSpeed=0.3 optiMoveAcceleration=0.09) tcp=t0_Flange; feature=Base
                    Waypoint WRHome: TCP in base x=651.404 y=-14.037 z=577.942 mm, rx=3.1416 ry=0 rz=0 rad; joints [-196.798, -95.185, 104.834, -99.59, -89.673, 73.253] deg; TCP offset x=0 y=0 z=0 mm, rx=0 ry=0 rz=3.1416 rad
                Script: Report(97)
            If Progress_run()
              Script: Report(50)
        Folder Buttons
          If In(ProgExe,[31,32,37,38,71,72,77,78])
            Script: Report(1)
            Folder AtHome?
              Timer (action=Reset) variable=T_Timeout
              Timer (action=Start) variable=T_Timeout
              Wait Condition expression=AtHomePos or (AtCenterPos and In(ProgExe,[71,72,77,78])) or T_Timeout>5
              If AtHomePos or (In(ProgExe,[71,72,77,78]) and AtCenterPos)
                'nop'
              Else 
                Script: Report(90)
            If Progress_run() and  not ((Di_SBR_L_X_Wp and ProgExe<50)  or (Di_SBR_R_X_Wp and ProgExe>50))
              Script: Report(92)
            If Progress_run()
              Folder Camera
                MoveJ speed 120 deg/s, acceleration 500 deg/s^2 (useActiveTCP=false positionType=JointAngles optimoveEnabled=false optiMoveSpeed=0.3 optiMoveAcceleration=0.09) tcp=t0_Flange; feature=Base
                  If In(ProgExe,[31,32])
                    SetCameraProg := 32
                    Waypoint WLBttnMidp: motionParameters(blendRadius=0.05); TCP in base x=-976.608 y=320.046 z=554.403 mm, rx=0 ry=3.1416 rz=0 rad; joints [-27.932, -58.226, 61.257, -92.971, -89.721, 62.073] deg
                    Waypoint WLCamLMB: TCP in base x=-1046.492 y=470.433 z=324.131 mm, rx=-0.2738 ry=3.1296 rz=0 rad; joints [-32.973, -41.135, 55.609, -104.414, -89.729, 47.088] deg
                  If In(ProgExe,[37,38])
                    SetCameraProg := 37
                    Waypoint WLBttnMidp: motionParameters(blendRadius=0.05); TCP in base x=-976.608 y=320.046 z=554.403 mm, rx=0 ry=3.1416 rz=0 rad; joints [-27.932, -58.226, 61.257, -92.971, -89.721, 62.073] deg
                    Waypoint WLCamLMB2: TCP in base x=-1046.492 y=576.368 z=294.652 mm, rx=-0.2738 ry=3.1296 rz=0 rad; joints [-37.258, -34.724, 46.673, -101.89, -89.735, 42.783] deg
                  If In(ProgExe,[71,72])
                    SetCameraProg := 72
                    Waypoint WpCenter: motionParameters(blendRadius=0.05); TCP in base x=-50 y=348.529 z=581.932 mm, rx=0 ry=3.1416 rz=0 rad; joints [-111.545, -128.858, 124.717, -85.8, -89.657, -21.591] deg; TCP offset x=0 y=0 z=0 mm, rx=0 ry=0 rz=3.1416 rad
                    Waypoint WRCamLMB: TCP in base x=-9.836 y=496.619 z=310.008 mm, rx=-0.2738 ry=3.1296 rz=0 rad; joints [-109.501, -99.356, 138.177, -128.761, -89.694, -29.281] deg; TCP offset x=0 y=0 z=0 mm, rx=0 ry=0 rz=3.1416 rad
                  If In(ProgExe,[77,78])
                    SetCameraProg := 77
                    Waypoint WpCenter: motionParameters(blendRadius=0.05); TCP in base x=-50 y=348.529 z=581.932 mm, rx=0 ry=3.1416 rz=0 rad; joints [-111.545, -128.858, 124.717, -85.8, -89.657, -21.591] deg; TCP offset x=0 y=0 z=0 mm, rx=0 ry=0 rz=3.1416 rad
                    Waypoint WRCamLMB2: TCP in base x=-9.836 y=605.743 z=283.054 mm, rx=-0.2738 ry=3.1296 rz=0 rad; joints [-105.879, -85.798, 129.08, -133.223, -89.721, -25.634] deg; TCP offset x=0 y=0 z=0 mm, rx=0 ry=0 rz=3.1416 rad
                Call CamAcquire
                Call CamCalculateCorectnPlane
            If Progress_run() and CamCorrectnOK≠ProgExe
              MoveL speed 1000 mm/s, acceleration 3000 mm/s^2 (useActiveTCP=false optimoveEnabled=false optiMoveSpeed=0.3 optiMoveAcceleration=0.09) tcp=t0_Flange; feature=Base
                If ProgExe<50
                  Waypoint WLBttnMidp: motionParameters(blendRadius=0.05); TCP in base x=-976.608 y=320.046 z=554.403 mm, rx=0 ry=3.1416 rz=0 rad; joints [-27.932, -58.226, 61.257, -92.971, -89.721, 62.073] deg
                  Waypoint WLHome: TCP in base x=-866.235 y=106.553 z=568.537 mm, rx=3.1416 ry=0 rz=0 rad; joints [-18.569, -73.864, 82.281, -98.358, -89.699, -108.526] deg
                Else 
                  Waypoint WpCenter: TCP in base x=-50 y=348.529 z=581.932 mm, rx=0 ry=3.1416 rz=0 rad; joints [-111.545, -128.858, 124.717, -85.8, -89.657, -21.591] deg; TCP offset x=0 y=0 z=0 mm, rx=0 ry=0 rz=3.1416 rad
                  STS_Reservation := 0
              Script: Report(91)
            If Progress_run()
              Folder Lumbar
                If In(ProgExe,[31,32,37,38,71,72,77,78])
                  Timer (action=Reset) variable=T_Timeout
                  Timer (action=Start) variable=T_Timeout
                  Script: Report(12)
                  Wait Condition expression=Flags[2] or T_Timeout>60 or DEBUG or Abort
                  If Flags[2] or DEBUG
                    MoveL speed 1000 mm/s, acceleration 3000 mm/s^2 (useActiveTCP=false optimoveEnabled=false optiMoveSpeed=0.3 optiMoveAcceleration=0.09) tcp=t4_Finger; feature=Base
                      Folder Press FW
                        If False
                          Waypoint WLLmbFw: TCP in base x=-785.023 y=519.426 z=306.838 mm, rx=-0.2738 ry=3.1296 rz=0 rad; joints [-39.124, -47.75, 61.996, -104.22, -89.71, 40.924] deg; TCP offset x=159 y=58 z=70 mm, rx=0 ry=0 rz=-3.1416 rad
                          Waypoint WLLmbFw2: TCP in base x=-787.926 y=626.666 z=276.111 mm, rx=-0.2738 ry=3.1296 rz=0 rad; joints [-43.172, -40.407, 52.022, -101.587, -89.716, 36.856] deg
                          Waypoint WRLmbFw: TCP in base x=217.007 y=523.124 z=293.128 mm, rx=-0.2738 ry=3.1296 rz=0 rad; joints [-113.579, -96.857, 129.584, -122.701, -89.677, -33.399] deg
                          Waypoint WRLmbFw2: TCP in base x=215.059 y=632.316 z=266.06 mm, rx=-0.2738 ry=3.1296 rz=0 rad; joints [-109.475, -84.368, 120.57, -126.176, -89.697, -29.275] deg
                        If In(ProgExe,[31,32])
                          Wp := pose_add(WLLmbFw,Base_w_correctn)
                        If In(ProgExe,[37,38])
                          Wp := pose_add(WLLmbFw2,Base_w_correctn)
                        If In(ProgExe,[71,72])
                          Wp := pose_add(WRLmbFw,Base_w_correctn)
                        If In(ProgExe,[77,78])
                          Wp := pose_add(WRLmbFw2,Base_w_correctn)
                        Waypoint Variable (Variable): variable=Wp
                        Force Frame feature=Joint_6_name; selection=[1, 0, 0, 0, 0, 0]; wrench=[-20, 10, -20, 0, 0, 0]; limitsForce=[0.05, 0.01, 0.05, 1.047198, 1.047198, 1.047198]; limitsMotion=[0.1, 0.1, 0.1, 0.349066, 0.349066, 0.349066]
                          Wait Sleep waitTime=0.7
                        ButtonPos := get_actual_tcp_pose()
                        Waypoint Variable (Variable): variable=Wp
                    Script: Report(3)
                  Else 
                    MoveJ speed 120 deg/s, acceleration 500 deg/s^2 (useActiveTCP=false positionType=JointAngles optimoveEnabled=false optiMoveSpeed=0.3 optiMoveAcceleration=0.09) tcp=t0_Flange; feature=Base
                      If ProgExe<50
                        Waypoint WLBttnMidp: motionParameters(blendRadius=0.05); TCP in base x=-976.608 y=320.046 z=554.403 mm, rx=0 ry=3.1416 rz=0 rad; joints [-27.932, -58.226, 61.257, -92.971, -89.721, 62.073] deg; TCP offset x=0 y=0 z=0 mm, rx=0 ry=0 rz=3.1416 rad
                        Waypoint WLHome: TCP in base x=-866.235 y=106.553 z=568.537 mm, rx=3.1416 ry=0 rz=0 rad; joints [-18.569, -73.864, 82.281, -98.358, -89.699, -108.526] deg
                      Else 
                        Waypoint WpCenter: TCP in base x=-50 y=348.529 z=581.932 mm, rx=0 ry=3.1416 rz=0 rad; joints [-111.545, -128.858, 124.717, -85.8, -89.657, -21.591] deg; TCP offset x=0 y=0 z=0 mm, rx=0 ry=0 rz=3.1416 rad
                        STS_Reservation := 0
                    Script: Report(95)
            If Progress_run()
              Folder Multiring
                If In(ProgExe,[32,38,72,78])
                  Timer (action=Reset) variable=T_Timeout
                  Timer (action=Start) variable=T_Timeout
                  Script: Report(11)
                  Wait Condition expression=Flags[1] or T_Timeout>60 or DEBUG or Abort
                  If Flags[1] or DEBUG
                    MoveL speed 1000 mm/s, acceleration 3000 mm/s^2 (useActiveTCP=false optimoveEnabled=false optiMoveSpeed=0.3 optiMoveAcceleration=0.09) tcp=t4_Finger; feature=Base
                      If False
                        Waypoint WLMultiringHi: TCP in base x=-766.371 y=505.747 z=321.008 mm, rx=-0.2738 ry=3.1296 rz=0 rad; joints [-39.188, -50.477, 65.229, -104.726, -89.708, 40.866] deg; TCP offset x=159 y=58 z=70 mm, rx=0 ry=0 rz=-3.1416 rad
                        Waypoint WLMultiringLo: TCP in base x=-766.487 y=502.365 z=299.18 mm, rx=-0.2738 ry=3.1296 rz=0 rad; joints [-39.045, -50.025, 66.731, -106.68, -89.708, 41.021] deg
                        Waypoint WLMultiringHi2: TCP in base x=-769.582 y=614.986 z=290.458 mm, rx=-0.2738 ry=3.1296 rz=0 rad; joints [-43.38, -43.245, 55.705, -102.432, -89.714, 36.656] deg
                        Waypoint WLMultiringLo2: TCP in base x=-767.873 y=608.483 z=269.439 mm, rx=-0.2738 ry=3.1296 rz=0 rad; joints [-43.2, -43.251, 57.884, -104.605, -89.713, 36.849] deg
                        Waypoint WRMultiringHi: TCP in base x=235.907 y=511.541 z=304.894 mm, rx=-0.2738 ry=3.1296 rz=0 rad; joints [-115.994, -98.646, 129.676, -121.005, -89.672, -35.825] deg
                        Waypoint WRMultiringLo: TCP in base x=235.896 y=508.024 z=287.162 mm, rx=-0.2738 ry=3.1296 rz=0 rad; joints [-116.168, -97.864, 131.14, -123.25, -89.677, -35.985] deg
                        Waypoint WRMultiringHi2: TCP in base x=234.761 y=620.702 z=278.623 mm, rx=-0.2738 ry=3.1296 rz=0 rad; joints [-111.505, -86.069, 120.908, -124.813, -89.693, -31.313] deg
                        Waypoint WRMultiringLo2: TCP in base x=235.553 y=618.433 z=259.689 mm, rx=-0.2738 ry=3.1296 rz=0 rad; joints [-111.65, -85.045, 122.127, -127.057, -89.699, -31.445] deg
                      Folder Press up
                        If ProgExe≟32
                          Wp0 := pose_add(WLMultiringLo,Base_w_correctn)
                        If ProgExe≟38
                          Wp0 := pose_add(WLMultiringLo2,Base_w_correctn)
                        If ProgExe≟72
                          Wp0 := pose_add(WRMultiringLo,Base_w_correctn)
                        If ProgExe≟78
                          Wp0 := pose_add(WRMultiringLo2,Base_w_correctn)
                        Wp0 := pose_trans(Wp0, p[0.02,0,0,0,0,0])
                        Wp := Wp0
                        Script: Wp[0]=ButtonPos[0]+0.01
                        Waypoint Variable (Variable): variable=Wp0
                        Waypoint Variable (Variable): variable=Wp
                        Set NoAction tcp=t4_Finger
                        Force Frame feature=Joint_6_name; selection=[0, 1, 1, 0, 0, 0]; wrench=[10, 20, -20, 0, 0, 0]; limitsForce=[0.01, 0.01, 0.025, 1.047198, 1.047198, 1.047198]; limitsMotion=[0.1, 0.1, 0.1, 0.349066, 0.349066, 0.349066]
                          Wait Sleep waitTime=1
                        Waypoint Variable (Variable): variable=Wp0
                      Folder Press down
                        If ProgExe≟32
                          Wp0 := pose_add(WLMultiringHi,Base_w_correctn)
                        If ProgExe≟38
                          Wp0 := pose_add(WLMultiringHi2,Base_w_correctn)
                        If ProgExe≟72
                          Wp0 := pose_add(WRMultiringHi,Base_w_correctn)
                        If ProgExe≟78
                          Wp0 := pose_add(WRMultiringHi2,Base_w_correctn)
                        Wp0 := pose_trans(Wp0, p[0.02,0,0,0,0,0])
                        Wp := Wp0
                        Script: Wp[0]=ButtonPos[0]+0.01
                        Waypoint Variable (Variable): variable=Wp0
                        Waypoint Variable (Variable): variable=Wp
                        Set NoAction tcp=t4_Finger
                        Force Frame feature=Joint_6_name; selection=[0, 1, 1, 0, 0, 0]; wrench=[10, 20, 20, 0, 0, 0]; limitsForce=[0.01, 0.01, 0.05, 1.047198, 1.047198, 1.047198]; limitsMotion=[0.1, 0.1, 0.1, 0.349066, 0.349066, 0.349066]
                          Wait Sleep waitTime=1
                        Waypoint Variable (Variable): variable=Wp0
                    Script: Report(2)
                  Else 
                    MoveJ speed 120 deg/s, acceleration 500 deg/s^2 (useActiveTCP=false positionType=JointAngles optimoveEnabled=false optiMoveSpeed=0.3 optiMoveAcceleration=0.09) tcp=t0_Flange; feature=Base
                      If ProgExe<50
                        Waypoint WLBttnMidp: motionParameters(blendRadius=0.05); TCP in base x=-976.608 y=320.046 z=554.403 mm, rx=0 ry=3.1416 rz=0 rad; joints [-27.932, -58.226, 61.257, -92.971, -89.721, 62.073] deg; TCP offset x=0 y=0 z=0 mm, rx=0 ry=0 rz=3.1416 rad
                        Waypoint WLHome: motionParameters(blendRadius=0.05); TCP in base x=-866.235 y=106.553 z=568.537 mm, rx=3.1416 ry=0 rz=0 rad; joints [-18.569, -73.864, 82.281, -98.358, -89.699, -108.526] deg
                      Else 
                        Waypoint WpCenter: TCP in base x=-50 y=348.529 z=581.932 mm, rx=0 ry=3.1416 rz=0 rad; joints [-111.545, -128.858, 124.717, -85.8, -89.657, -21.591] deg; TCP offset x=0 y=0 z=0 mm, rx=0 ry=0 rz=3.1416 rad
                        STS_Reservation := 0
                    Script: Report(95)
            If Progress_run()
              MoveJ speed 120 deg/s, acceleration 500 deg/s^2 (useActiveTCP=false positionType=JointAngles optimoveEnabled=false optiMoveSpeed=0.3 optiMoveAcceleration=0.09) tcp=t0_Flange; feature=Base
                If ProgExe<50
                  Waypoint WLBttnMidp: TCP in base x=-976.608 y=320.046 z=554.403 mm, rx=0 ry=3.1416 rz=0 rad; joints [-27.932, -58.226, 61.257, -92.971, -89.721, 62.073] deg; TCP offset x=0 y=0 z=0 mm, rx=0 ry=0 rz=3.1416 rad
                  Waypoint WLHome: TCP in base x=-866.235 y=106.553 z=568.537 mm, rx=3.1416 ry=0 rz=0 rad; joints [-18.569, -73.864, 82.281, -98.358, -89.699, -108.526] deg
                Else 
                  Waypoint WpCenter: TCP in base x=-50 y=348.529 z=581.932 mm, rx=0 ry=3.1416 rz=0 rad; joints [-111.545, -128.858, 124.717, -85.8, -89.657, -21.591] deg; TCP offset x=0 y=0 z=0 mm, rx=0 ry=0 rz=3.1416 rad
                  STS_Reservation := 0
              Script: Report(50)
        Folder Program finished
          ProgDn := ProgExe
          ProgExe := 0
      Folder Parking
        If Parking≟10 or ProgExe≟1010
          Wait Condition expression=EvtDock≤0
          If AtLHomePos
            MoveJ speed 120 deg/s, acceleration 500 deg/s^2 (useActiveTCP=true positionType=JointAngles optimoveEnabled=false optiMoveSpeed=0.3 optiMoveAcceleration=0.09) feature=Base
              Waypoint WLHome0: motionParameters(blendRadius=0.1); TCP in base x=-460.734 y=106.553 z=568.537 mm, rx=-2.2214 ry=2.2214 rz=0 rad; joints [-34.699, -114.011, 119.5, -95.429, -89.656, -34.68] deg; TCP offset x=0 y=0 z=0 mm, rx=0 ry=0 rz=3.1416 rad
              Waypoint WpCenter: TCP in base x=-50 y=348.529 z=581.932 mm, rx=0 ry=3.1416 rz=0 rad; joints [-111.545, -128.858, 124.717, -85.8, -89.657, -21.591] deg; TCP offset x=0 y=0 z=0 mm, rx=0 ry=0 rz=3.1416 rad
          If AtRHomePos
            MoveJ speed 120 deg/s, acceleration 500 deg/s^2 (useActiveTCP=false positionType=JointAngles optimoveEnabled=false optiMoveSpeed=0.3 optiMoveAcceleration=0.09) tcp=t0_Flange; feature=Base
              Waypoint WpCenter: TCP in base x=-50 y=348.529 z=581.932 mm, rx=0 ry=3.1416 rz=0 rad; joints [-111.545, -128.858, 124.717, -85.8, -89.657, -21.591] deg
          Parking := 0
          If DEBUG
            ProgExe := 0
        If Parking≟11 or ProgExe≟1011
          Wait Condition expression=EvtDock≤0
          If AtLHomePos
            MoveJ speed 120 deg/s, acceleration 500 deg/s^2 (useActiveTCP=true positionType=JointAngles optimoveEnabled=false optiMoveSpeed=0.3 optiMoveAcceleration=0.09) feature=Base
              Waypoint WLHome0: motionParameters(blendRadius=0.05); TCP in base x=-460.734 y=106.553 z=568.537 mm, rx=-2.2214 ry=2.2214 rz=0 rad; joints [-34.699, -114.011, 119.5, -95.429, -89.656, -34.68] deg; TCP offset x=0 y=0 z=0 mm, rx=0 ry=0 rz=3.1416 rad
              Waypoint WpCenter: motionParameters(blendRadius=0.1); TCP in base x=-50 y=348.529 z=581.932 mm, rx=0 ry=3.1416 rz=0 rad; joints [-111.545, -128.858, 124.717, -85.8, -89.657, -21.591] deg; TCP offset x=0 y=0 z=0 mm, rx=0 ry=0 rz=3.1416 rad
              Waypoint WpPark0: motionParameters(blendRadius=0.1); TCP in base x=-173.588 y=120.798 z=947.577 mm, rx=-2.2245 ry=-2.2153 rz=0.001 rad; joints [-90.355, -130.078, 83.552, -43.476, -89.706, 89.65] deg; TCP offset x=0 y=0 z=0 mm, rx=0 ry=0 rz=3.1416 rad
              Waypoint WpPark1: motionParameters(blendRadius=0.05); TCP in base x=121.203 y=255.21 z=1195.147 mm, rx=-1.7636 ry=-1.7554 rz=-0.7332 rad; joints [-180.212, -111.325, 44.19, -22.632, -44.842, -0.325] deg
              Waypoint WpPark: TCP in base x=121.203 y=255.21 z=1282.913 mm, rx=-1.7636 ry=-1.7554 rz=-0.7332 rad; joints [-180, -89.998, -0.001, 0.001, -45, 0] deg
          If AtRHomePos
            MoveJ speed 120 deg/s, acceleration 500 deg/s^2 (useActiveTCP=false positionType=JointAngles optimoveEnabled=false optiMoveSpeed=0.3 optiMoveAcceleration=0.09) tcp=t0_Flange; feature=Base
              Waypoint WpCenter: motionParameters(blendRadius=0.1); TCP in base x=-50 y=348.529 z=581.932 mm, rx=0 ry=3.1416 rz=0 rad; joints [-111.545, -128.858, 124.717, -85.8, -89.657, -21.591] deg; TCP offset x=0 y=0 z=0 mm, rx=0 ry=0 rz=3.1416 rad
              Waypoint WpPark0: motionParameters(blendRadius=0.1); TCP in base x=-173.588 y=120.798 z=947.577 mm, rx=-2.2245 ry=-2.2153 rz=0.001 rad; joints [-90.355, -130.078, 83.552, -43.476, -89.706, 89.65] deg; TCP offset x=0 y=0 z=0 mm, rx=0 ry=0 rz=3.1416 rad
              Waypoint WpPark1: motionParameters(blendRadius=0.05); TCP in base x=121.203 y=255.21 z=1195.147 mm, rx=-1.7636 ry=-1.7554 rz=-0.7332 rad; joints [-180.212, -111.325, 44.19, -22.632, -44.842, -0.325] deg
              Waypoint WpPark: TCP in base x=121.203 y=255.21 z=1282.913 mm, rx=-1.7636 ry=-1.7554 rz=-0.7332 rad; joints [-180, -89.998, -0.001, 0.001, -45, 0] deg
          If AtCenterPos
            MoveJ speed 120 deg/s, acceleration 500 deg/s^2 (useActiveTCP=false positionType=JointAngles optimoveEnabled=false optiMoveSpeed=0.3 optiMoveAcceleration=0.09) tcp=t0_Flange; feature=Base
              Waypoint WpPark0: motionParameters(blendRadius=0.1); TCP in base x=-173.588 y=120.798 z=947.577 mm, rx=-2.2245 ry=-2.2153 rz=0.001 rad; joints [-90.355, -130.078, 83.552, -43.476, -89.706, 89.65] deg
              Waypoint WpPark1: motionParameters(blendRadius=0.05); TCP in base x=121.203 y=255.21 z=1195.147 mm, rx=-1.7636 ry=-1.7554 rz=-0.7332 rad; joints [-180.212, -111.325, 44.19, -22.632, -44.842, -0.325] deg
              Waypoint WpPark: TCP in base x=121.203 y=255.21 z=1282.913 mm, rx=-1.7636 ry=-1.7554 rz=-0.7332 rad; joints [-180, -89.998, -0.001, 0.001, -45, 0] deg
          Parking := 0
          If DEBUG
            ProgExe := 0
        If Parking≟1 or ProgExe≟1001
          If AtParkPos
            MoveJ speed 120 deg/s, acceleration 500 deg/s^2 (useActiveTCP=false positionType=JointAngles optimoveEnabled=false optiMoveSpeed=0.3 optiMoveAcceleration=0.09) tcp=t0_Flange; feature=Base
              Waypoint WpPark1: motionParameters(blendRadius=0.05); TCP in base x=121.203 y=255.21 z=1195.147 mm, rx=-1.7636 ry=-1.7554 rz=-0.7332 rad; joints [-180.212, -111.325, 44.19, -22.632, -44.842, -0.325] deg
              Waypoint WpPark0: motionParameters(blendRadius=0.1); TCP in base x=-173.588 y=120.798 z=947.577 mm, rx=-2.2245 ry=-2.2153 rz=0.001 rad; joints [-90.355, -130.078, 83.552, -43.476, -89.706, 89.65] deg
              Waypoint WpCenter: motionParameters(blendRadius=0.05); TCP in base x=-50 y=348.529 z=581.932 mm, rx=0 ry=3.1416 rz=0 rad; joints [-111.545, -128.858, 124.717, -85.8, -89.657, -21.591] deg; TCP offset x=0 y=0 z=0 mm, rx=0 ry=0 rz=3.1416 rad
              Waypoint WLHome0: motionParameters(blendRadius=0.05); TCP in base x=-460.734 y=106.553 z=568.537 mm, rx=-2.2214 ry=2.2214 rz=0 rad; joints [-34.699, -114.011, 119.5, -95.429, -89.656, -34.68] deg; TCP offset x=0 y=0 z=0 mm, rx=0 ry=0 rz=3.1416 rad
              Waypoint WLHome: TCP in base x=-866.235 y=106.553 z=568.537 mm, rx=3.1416 ry=0 rz=0 rad; joints [-18.569, -73.864, 82.281, -98.358, -89.699, -108.526] deg
              STS_Reservation := 1
          If AtCenterPos
            MoveJ speed 120 deg/s, acceleration 500 deg/s^2 (useActiveTCP=false positionType=JointAngles optimoveEnabled=false optiMoveSpeed=0.3 optiMoveAcceleration=0.09) tcp=t0_Flange; feature=Base
              Waypoint WLHome0: motionParameters(blendRadius=0.05); TCP in base x=-460.734 y=106.553 z=568.537 mm, rx=-2.2214 ry=2.2214 rz=0 rad; joints [-34.699, -114.011, 119.5, -95.429, -89.656, -34.68] deg
              Waypoint WLHome referenceName=WLHome: TCP in base x=-866.235 y=106.553 z=568.537 mm, rx=3.1416 ry=0 rz=0 rad; joints [-18.569, -73.864, 82.281, -98.358, -89.699, -108.526] deg
              STS_Reservation := 1
          If AtRHomePos
            MoveJ speed 120 deg/s, acceleration 500 deg/s^2 (useActiveTCP=false positionType=JointAngles optimoveEnabled=false optiMoveSpeed=0.3 optiMoveAcceleration=0.09) tcp=t0_Flange; feature=Base
              Waypoint WpCenter: motionParameters(blendRadius=0.05); TCP in base x=-50 y=348.529 z=581.932 mm, rx=0 ry=3.1416 rz=0 rad; joints [-111.545, -128.858, 124.717, -85.8, -89.657, -21.591] deg; TCP offset x=0 y=0 z=0 mm, rx=0 ry=0 rz=3.1416 rad
              Waypoint WLHome0: motionParameters(blendRadius=0.05); TCP in base x=-460.734 y=106.553 z=568.537 mm, rx=-2.2214 ry=2.2214 rz=0 rad; joints [-34.699, -114.011, 119.5, -95.429, -89.656, -34.68] deg; TCP offset x=0 y=0 z=0 mm, rx=0 ry=0 rz=3.1416 rad
              Waypoint WLHome: TCP in base x=-866.235 y=106.553 z=568.537 mm, rx=3.1416 ry=0 rz=0 rad; joints [-18.569, -73.864, 82.281, -98.358, -89.699, -108.526] deg
              STS_Reservation := 1
          Parking := 0
          If DEBUG
            ProgExe := 0
        If Parking≟2 or ProgExe≟1002
          If AtParkPos
            MoveJ speed 120 deg/s, acceleration 500 deg/s^2 (useActiveTCP=false positionType=JointAngles optimoveEnabled=false optiMoveSpeed=0.3 optiMoveAcceleration=0.09) tcp=t0_Flange; feature=Base
              Waypoint WpPark1: motionParameters(blendRadius=0.05); TCP in base x=121.203 y=255.21 z=1195.147 mm, rx=-1.7636 ry=-1.7554 rz=-0.7332 rad; joints [-180.212, -111.325, 44.19, -22.632, -44.842, -0.325] deg
              Waypoint WpPark0: motionParameters(blendRadius=0.1); TCP in base x=-173.588 y=120.798 z=947.577 mm, rx=-2.2245 ry=-2.2153 rz=0.001 rad; joints [-90.355, -130.078, 83.552, -43.476, -89.706, 89.65] deg
              Waypoint WpCenter: motionParameters(blendRadius=0.091); TCP in base x=-50 y=348.529 z=581.932 mm, rx=0 ry=3.1416 rz=0 rad; joints [-111.545, -128.858, 124.717, -85.8, -89.657, -21.591] deg; TCP offset x=0 y=0 z=0 mm, rx=0 ry=0 rz=3.1416 rad
              Waypoint WRHome: TCP in base x=651.404 y=-14.037 z=577.942 mm, rx=3.1416 ry=0 rz=0 rad; joints [-196.798, -95.185, 104.834, -99.59, -89.673, 73.253] deg; TCP offset x=0 y=0 z=0 mm, rx=0 ry=0 rz=3.1416 rad
              STS_Reservation := 2
          If AtCenterPos
            MoveJ speed 120 deg/s, acceleration 500 deg/s^2 (useActiveTCP=true positionType=JointAngles optimoveEnabled=false optiMoveSpeed=0.3 optiMoveAcceleration=0.09) feature=Base
              Waypoint WRHome: TCP in base x=651.404 y=-14.037 z=577.942 mm, rx=3.1416 ry=0 rz=0 rad; joints [-196.798, -95.185, 104.834, -99.59, -89.673, 73.253] deg
              STS_Reservation := 2
          If AtLHomePos
            MoveJ speed 120 deg/s, acceleration 500 deg/s^2 (useActiveTCP=false positionType=JointAngles optimoveEnabled=false optiMoveSpeed=0.3 optiMoveAcceleration=0.09) tcp=t0_Flange; feature=Base
              Waypoint WLHome0: motionParameters(blendRadius=0.05); TCP in base x=-460.734 y=106.553 z=568.537 mm, rx=-2.2214 ry=2.2214 rz=0 rad; joints [-34.699, -114.011, 119.5, -95.429, -89.656, -34.68] deg
              Waypoint WpCenter: motionParameters(blendRadius=0.1); TCP in base x=-50 y=348.529 z=581.932 mm, rx=0 ry=3.1416 rz=0 rad; joints [-111.545, -128.858, 124.717, -85.8, -89.657, -21.591] deg; TCP offset x=0 y=0 z=0 mm, rx=0 ry=0 rz=3.1416 rad
              Waypoint WRHome: TCP in base x=651.404 y=-14.037 z=577.942 mm, rx=3.1416 ry=0 rz=0 rad; joints [-196.798, -95.185, 104.834, -99.59, -89.673, 73.253] deg; TCP offset x=0 y=0 z=0 mm, rx=0 ry=0 rz=3.1416 rad
              STS_Reservation := 2
          Parking := 0
          If DEBUG
            ProgExe := 0
Thread Thread_1 (runOnlyOnce=false)
  Folder Continuous calculations
    Folder get live force and tcp pos
      P_act := get_actual_tcp_pose()
      V_act := get_actual_tcp_speed()
      V_act_norm := norm(V_act)
      P_Flange := get_actual_tool_flange_pose()
      D_rel := pose_sub(P_act, P_ini)
      Folder Detect home positions
        AtLHomePos := PosDist(P_Flange, WLHome)<0.005
        AtRHomePos := PosDist(P_Flange, WRHome)<0.005
        AtCenterPos := PosDist(P_Flange, WpCenter)<0.005
        AtParkPos := PosDist(P_Flange, WpPark)<0.005
        If InRange(ProgExe,10,49)
          AtHomePos := AtLHomePos
        ElseIf InRange(ProgExe,50,89)
          AtHomePos := AtRHomePos
        Else 
          AtHomePos := AtLHomePos or AtRHomePos
      Folder Detect docking signal
        If P_Flange[0]<0
          AdapterDocked := Di_Docked_L
        Else 
          AdapterDocked := Di_Docked_R
      Folder Calculate actual offset in tool frame
        If ProgExe≟15
          TempWp := pose_sub(WLBuckleSpa1,Base_w_correctn)
          BklToolDist := pose_trans(pose_inv(TempWp), P_act)
        If ProgExe≟16
          TempWp := pose_sub(WLBuckleSpa3,Base_w_correctn)
          BklToolDist := pose_trans(pose_inv(TempWp), P_act)
        If ProgExe≟55
          TempWp := pose_sub(WRBuckleSpa1,Base_w_correctn)
          BklToolDist := pose_trans(pose_inv(TempWp), P_act)
        If ProgExe≟56
          TempWp := pose_sub(WRBuckleSpa3,Base_w_correctn)
          BklToolDist := pose_trans(pose_inv(TempWp), P_act)
      Folder InterlockOutput
        If P_Flange[1]<0.45
          Set DigitalOutput pin=Do_SafePosition; digitalValue=1
        ElseIf P_Flange[0]>0.65
          Set DigitalOutput pin=Do_SafePosition; digitalValue=1
        ElseIf InRange(P_Flange[0],-0.35,0)
          Set DigitalOutput pin=Do_SafePosition; digitalValue=1
        Else 
          Set DigitalOutput pin=Do_SafePosition; digitalValue=0
    Folder Modbus mapping
      Folder Heartbeat
        Timer (action=Start) variable(name=T_Heartbeat)
        If T_Heartbeat≥1
          Timer (action=Reset) variable=T_Heartbeat
          If STS_Heartbeat
            STS_Heartbeat := False
          Else 
            STS_Heartbeat := True
      Folder Safe position
        Folder L
          STS_Safe_i1 := True
          If pose_dist(P_act, WLConnSpa1)<0.08
            STS_Safe_i1 := False
          If pose_dist(P_act, WLUnplug1_3)<0.05
            STS_Safe_i1 := False
          If pose_dist(P_act, WLBuckleSpa1)<0.2
            STS_Safe_i1 := False
          If pose_dist(P_act, WLLmbFw)<0.05
            STS_Safe_i1 := False
          If pose_dist(P_act, WLLmbFw2)<0.05
            STS_Safe_i1 := False
        Folder R
          STS_Safe_i2 := True
          If pose_dist(P_act, WRConnSpa1)<0.08
            STS_Safe_i2 := False
          If pose_dist(P_act, WRUnpgSpa1_3)<0.05
            STS_Safe_i2 := False
          If pose_dist(P_act, WRBuckleSpa1)<0.2
            STS_Safe_i2 := False
          If pose_dist(P_act, WRLmbFw)<0.05
            STS_Safe_i2 := False
          If pose_dist(P_act, WRLmbFw2)<0.05
            STS_Safe_i2 := False
      Folder Outputs
        Script: write_port_register(129,STS_Progress)
        Script: write_port_register(131,STS_Reservation)
        Script: write_port_register(134,binary_list_to_integer([Di_Docked_L,Di_Docked_R,NormalMode,STS_Heartbeat,STS_Safe_i1,STS_Safe_i2]))
      Folder Inputs
        CMD_Reserve_i1 := read_port_register(160)
        CMD_Reserve_i2 := read_port_register(161)
        CMD_Timeout_i1 := read_port_register(162)
        CMD_Timeout_i2 := read_port_register(163)
        CMD_Program_i1 := read_port_register(164)
        CMD_Program_i2 := read_port_register(165)
        CMD_Flags_i1 := read_port_register(170)
        CMD_Flags_i2 := read_port_register(171)
        CMD_Heartbt_i1 := read_port_register(180)
        CMD_Heartbt_i2 := read_port_register(181)
      Folder Generate flags
        Flags_i1 := integer_to_binary_list(CMD_Flags_i1)
        Flags_i2 := integer_to_binary_list(CMD_Flags_i2)
        If InRange(ProgExe,10,49)
          Flags := Flags_i1
        ElseIf InRange(ProgExe,50,89)
          Flags := Flags_i2
    Folder Operator call deactivation
      If Do_Blue or Do_Horn
        Timer (action=Start) variable(name=T_Call)
        If not  NormalMode and T_Call>4
          Set DigitalOutput pin=Do_Blue; digitalValue=0
          Set DigitalOutput pin=Do_Horn; digitalValue=0
          Mute := True
      Else 
        Timer (action=Stop) variable=T_Call
        Timer (action=Reset) variable=T_Call
      If ProgExe>0
        Mute := False
    Folder Abort
      If Flags_i1[14] and (InRange(ProgExe,10,49) or AdapterReady_L)
        Abort := True
      ElseIf Flags_i2[14] and (InRange(ProgExe,50,89) or AdapterReady_R)
        Abort := True
      If AtHomePos or AtCenterPos
        Abort := False
      If Abort
        If AdapterReady_L or AdapterReady_R
          EvtDock := 1
    Folder Speed
      Timer (action=Start) variable(name=T_SpeedSet)
      If T_SpeedSet>2 and  not DEBUG
        Script: socket_send_string("set speed")
        SuppressedNode
          Script: socket_send_string(0.9)
        Script: socket_send_string(1.0)
        Script: socket_send_byte(10)
        Timer (action=Reset) variable=T_SpeedSet
    Wait Sleep waitTime=0.01
  Folder ReservationControl
    'Request reservation, disconnect preference'
    If STS_Reservation≟0 and ProgExe≟0 and Parking≟0
      If CMD_Reserve_i1≟1 and In(CMD_Program_i1,[21,22,23])
        'request reservation'
        If AtLHomePos or AdapterReady_L
          STS_Reservation := 1
        Else 
          Parking := 1
      If CMD_Reserve_i2≟2 and In(CMD_Program_i2,[61,62,63])
        'request reservation'
        If AtRHomePos or AdapterReady_R
          STS_Reservation := 2
        Else 
          Parking := 2
      If CMD_Reserve_i1≟1
        'request reservation'
        If AtLHomePos or AdapterReady_L
          STS_Reservation := 1
        ElseIf In(CMD_Program_i1,[15,16])
          'Special case to save time when moving to buckle'
          If AtCenterPos
            STS_Reservation := 1
          Else 
            Parking := 10
        Else 
          Parking := 1
      If CMD_Reserve_i2≟2
        'request reservation'
        If AtRHomePos or AdapterReady_R
          STS_Reservation := 2
        ElseIf In(CMD_Program_i2,[71,72,77,78])
          'Special case to save time when moving to buttons'
          If AtCenterPos
            STS_Reservation := 2
          Else 
            Parking := 10
        Else 
          Parking := 2
    'Timeout reservation - station keeps reservation for a while to prevent other app stealing the process'
    'Timeout is configurable, so application can control how long to keep robot before letting other app'
    If STS_Progress≟0 and STS_Reservation≠0 and Parking≟0
      If STS_Reservation≟1 and CMD_Reserve_i1≟1
        'nop'
      ElseIf STS_Reservation≟2 and CMD_Reserve_i2≟2
        'nop'
      Else 
        If STS_Reservation≟1
          T_KeepReservtn := CMD_Timeout_i1
        If STS_Reservation≟2
          T_KeepReservtn := CMD_Timeout_i2
        Timer (action=Start) variable(name=T_Unreserve)
        If T_Unreserve>T_KeepReservtn
          STS_Reservation := 0
    Else 
      Timer (action=Stop) variable=T_Unreserve
      Timer (action=Reset) variable=T_Unreserve
    'Force release reservation from app - in case of intervetion'
    If STS_Reservation≟0 and STS_Progress≟0 and  not DEBUG
      If In(CMD_Reserve_i1,[98,99]) and  not In(CMD_Reserve_i2,[98,99]) and  not AtParkPos
        If AtRHomePos
          STS_Reservation := 2
        Else 
          Parking := 2
      If In(CMD_Reserve_i2,[98,99]) and  not In(CMD_Reserve_i1,[98,99]) and  not AtParkPos
        If AtLHomePos
          STS_Reservation := 1
        Else 
          Parking := 1
      If In(CMD_Reserve_i1,[98,99]) and In(CMD_Reserve_i2,[98,99])
        If AtParkPos
          STS_Reservation := 0
        Else 
          Parking := 11
      If (CMD_Reserve_i1≟99 or CMD_Reserve_i2≟99) and  not Mute
        Set DigitalOutput pin=Do_Blue; digitalValue=1
        Set DigitalOutput pin=Do_Horn; digitalValue=1
  Folder Program control
    'Start new Prog / Confirm Prog Running'
    If STS_Progress≟0 and ProgExe≟0  and  not Abort and  not DEBUG
      If InRange(CMD_Program_i1,10,49) and STS_Reservation≟1
        ProgExe := CMD_Program_i1
        T_KeepReservtn := CMD_Timeout_i1
        Script: Report(0)
      If InRange(CMD_Program_i2,50,89) and STS_Reservation≟2
        ProgExe := CMD_Program_i2
        T_KeepReservtn := CMD_Timeout_i2
        Script: Report(0)
    'Ack results - get ready for new prg'
    If ProgExe≟0 and Progress_finished()
      If InRange(ProgDn,10,49) and CMD_Program_i1≠ProgDn
        STS_Progress := 0
        If In(CMD_Program_i1,[21,22,23]) or In(CMD_Program_i2,[61,62,63])
          'unplug preference - unreserve immediatelly'
          STS_Reservation := 0
      If InRange(ProgDn,50,89) and CMD_Program_i2≠ProgDn
        STS_Progress := 0
        If In(CMD_Program_i1,[21,22,23]) or In(CMD_Program_i2,[61,62,63])
          'unplug preference - unreserve immediatelly'
          STS_Reservation := 0
SubProgram WaitForNormalMode [hidden by the author, left out]
SubProgram  [hidden by the author, left out]
SubProgram  [hidden by the author, left out]
SubProgram  [hidden by the author, left out]
SubProgram  [hidden by the author, left out]
Event  expression=SetCameraProg>0
  Folder Set program to camera in advance
    Set DigitalOutput pin=CnxDO_Trig; digitalValue=0
    Set DigitalOutput pin=CnxDO_TrigEn; digitalValue=1
    Script: modbus_delete_signal("CnxAO_Program")
    Script: modbus_add_signal("10.142.142.43", 255, 2001, 16, "CnxAO_Program", True ,1)
    Script: modbus_set_output_register("CnxAO_Program",SetCameraProg, False )
    Wait Sleep waitTime=0.2
    Set DigitalOutput pin=CnxDO_SetUsrDta; digitalValue=1
    Wait DigitalInput pin=CnxDi_UsrDtaAck; digitalValue=1
    Set DigitalOutput pin=CnxDO_SetUsrDta; digitalValue=0
    Set DigitalOutput pin=CnxDO_SoftEvt0; digitalValue=1
    Wait DigitalInput pin=CnxDI_Evt0Ack; digitalValue=1
    Set DigitalOutput pin=CnxDO_SoftEvt0; digitalValue=0
    Timer (action=Reset) variable=CamTimeout
    Timer (action=Start) variable=CamTimeout
    Wait Condition expression=CnxAI_Program≟SetCameraProg or CamTimeout>3
    If CnxAI_Program≠SetCameraProg
      Script: textmsg("set cam prog failed, trying trigger")
      Folder For the first time it needs trigger when going online
        Set DigitalOutput pin=CnxDO_Trig; digitalValue=1
        Wait Sleep waitTime=1
        Set DigitalOutput pin=CnxDO_Trig; digitalValue=0
      If CnxAI_Program≠SetCameraProg
        SuppressedNode
          Popup Error (haltProgram=false message=Error: camera program not set inputType=Text)
      Else 
        Wait Sleep waitTime=0.5
        SetCameraProg := 0
    Else 
      Wait Sleep waitTime=0.5
      SetCameraProg := 0
  If SetCameraProg>0
    'repeat on fail'
    Wait Sleep waitTime=3
    Folder Set program to camera in advance
      Set DigitalOutput pin=CnxDO_Trig; digitalValue=0
      Set DigitalOutput pin=CnxDO_TrigEn; digitalValue=1
      Script: modbus_delete_signal("CnxAO_Program")
      Script: modbus_add_signal("10.142.142.43", 255, 2001, 16, "CnxAO_Program", True ,1)
      Script: modbus_set_output_register("CnxAO_Program",SetCameraProg, False )
      Wait Sleep waitTime=0.2
      Set DigitalOutput pin=CnxDO_SetUsrDta; digitalValue=1
      Wait DigitalInput pin=CnxDi_UsrDtaAck; digitalValue=1
      Set DigitalOutput pin=CnxDO_SetUsrDta; digitalValue=0
      Set DigitalOutput pin=CnxDO_SoftEvt0; digitalValue=1
      Wait DigitalInput pin=CnxDI_Evt0Ack; digitalValue=1
      Set DigitalOutput pin=CnxDO_SoftEvt0; digitalValue=0
      Timer (action=Reset) variable=CamTimeout
      Timer (action=Start) variable=CamTimeout
      Wait Condition expression=CnxAI_Program≟SetCameraProg or CamTimeout>3
      If CnxAI_Program≠SetCameraProg
        Script: textmsg("set cam prog failed, trying trigger")
        Folder For the first time it needs trigger when going online
          Set DigitalOutput pin=CnxDO_Trig; digitalValue=1
          Wait Sleep waitTime=1
          Set DigitalOutput pin=CnxDO_Trig; digitalValue=0
        If CnxAI_Program≠SetCameraProg
          SuppressedNode
            Popup Error (haltProgram=false message=Error: camera program not set inputType=Text)
        Else 
          Wait Sleep waitTime=0.5
          SetCameraProg := 0
      Else 
        Wait Sleep waitTime=0.5
        SetCameraProg := 0
  If SetCameraProg>0
    'repeat on fail'
    Wait Sleep waitTime=3
    Folder Set program to camera in advance
      Set DigitalOutput pin=CnxDO_Trig; digitalValue=0
      Set DigitalOutput pin=CnxDO_TrigEn; digitalValue=1
      Script: modbus_delete_signal("CnxAO_Program")
      Script: modbus_add_signal("10.142.142.43", 255, 2001, 16, "CnxAO_Program", True ,1)
      Script: modbus_set_output_register("CnxAO_Program",SetCameraProg, False )
      Wait Sleep waitTime=0.2
      Set DigitalOutput pin=CnxDO_SetUsrDta; digitalValue=1
      Wait DigitalInput pin=CnxDi_UsrDtaAck; digitalValue=1
      Set DigitalOutput pin=CnxDO_SetUsrDta; digitalValue=0
      Set DigitalOutput pin=CnxDO_SoftEvt0; digitalValue=1
      Wait DigitalInput pin=CnxDI_Evt0Ack; digitalValue=1
      Set DigitalOutput pin=CnxDO_SoftEvt0; digitalValue=0
      Timer (action=Reset) variable=CamTimeout
      Timer (action=Start) variable=CamTimeout
      Wait Condition expression=CnxAI_Program≟SetCameraProg or CamTimeout>3
      If CnxAI_Program≠SetCameraProg
        Script: textmsg("set cam prog failed, trying trigger")
        Folder For the first time it needs trigger when going online
          Set DigitalOutput pin=CnxDO_Trig; digitalValue=1
          Wait Sleep waitTime=1
          Set DigitalOutput pin=CnxDO_Trig; digitalValue=0
        If CnxAI_Program≠SetCameraProg
          SuppressedNode
            Popup Error (haltProgram=false message=Error: camera program not set inputType=Text)
        Else 
          Wait Sleep waitTime=0.5
          SetCameraProg := 0
      Else 
        Wait Sleep waitTime=0.5
        SetCameraProg := 0
  If SetCameraProg>0
    Popup Error (haltProgram=false message=Error: camera program not set inputType=Text)
SubProgram -> CamAcquire
SubProgram -> CamCalculateCorectnPlane
Event  expression=EvtDock>0
  Folder Dock
    MoveL speed 1000 mm/s, acceleration 3000 mm/s^2 (useActiveTCP=false optimoveEnabled=false optiMoveSpeed=0.3 optiMoveAcceleration=0.09) tcp=t2_Gripper; feature=Base
      If EvtDock≟2
        Folder Force mvts
          Set NoAction tcp=t2_Gripper
          Wp0 := P_act
          Force Frame feature=Joint_6_name; selection=[0, 1, 0, 0, 0, 0]; wrench=[0, -20, 0, 0, 0, 0]; limitsForce=[0.15, 0.1, 0.15, 1.047198, 1.047198, 1.047198]; limitsMotion=[0.1, 0.1, 0.1, 0.349066, 0.349066, 0.349066]
            Wait Sleep waitTime=1
          Force Frame feature=Joint_6_name; selection=[1, 0, 1, 1, 0, 0]; wrench=[0, -10, 0, 0, 0, 0]; limitsForce=[0.15, 0.05, 0.1, 1.047198, 1.047198, 1.047198]; limitsMotion=[0.1, 0.1, 0.1, 0.349066, 0.349066, 0.349066]
            Wait Sleep waitTime=0.2
            Call GripperClose
            Wait Sleep waitTime=0.2
          If T_Gripper>3
            Call GripperOpen
            MoveL speed 500 mm/s, acceleration 1200 mm/s^2 (useActiveTCP=true optimoveEnabled=false optiMoveSpeed=0.3 optiMoveAcceleration=0.09) feature=Base
              Waypoint Variable (Variable): variable=Wp0
            Force Frame feature=Joint_6_name; selection=[0, 1, 0, 0, 0, 0]; wrench=[0, -20, 0, 0, 0, 0]; limitsForce=[0.15, 0.1, 0.15, 1.047198, 1.047198, 1.047198]; limitsMotion=[0.1, 0.1, 0.1, 0.349066, 0.349066, 0.349066]
              Wait Sleep waitTime=1
            Force Frame feature=Joint_6_name; selection=[1, 0, 1, 0, 0, 0]; wrench=[0, -10, 0, 0, 0, 0]; limitsForce=[0.15, 0.05, 0.1, 1.047198, 1.047198, 1.047198]; limitsMotion=[0.1, 0.1, 0.1, 0.349066, 0.349066, 0.349066]
              Wait Sleep waitTime=0.2
              Call GripperClose
              Wait Sleep waitTime=0.2
          If T_Gripper>3
            Call GripperOpen
            MoveL speed 500 mm/s, acceleration 1200 mm/s^2 (useActiveTCP=true optimoveEnabled=false optiMoveSpeed=0.3 optiMoveAcceleration=0.09) feature=Base
              Waypoint Variable (Variable): variable=Wp0
              EvtDock := -97
          If EvtDock≟2
            MoveDirectionNode (selectedDirection=YPlus) feature=Joint_6_name
              Until DISTANCE (allowActions=false deceleration=3 distanceNodeType=BLEND) Distance=0.1; motionParameters(blendRadius=0.05)
      If InRange(EvtDock,1,2)
        If P_Flange[0]<0
          WpDock := WLDock
          WpHome := WLHome
        Else 
          WpDock := WRDock
          WpHome := WRHome
        Script: Report(40)
        Wp := pose_trans(WpDock, p[0,0.25,0,0,0,0])
        Waypoint Variable (Variable): motionParameters(blendRadius=0.05); variable=Wp
        Waypoint Variable (Variable): variable=WpDock
        Call GripperOpen
        Waypoint Variable (Variable): variable=Wp
        MoveL speed 1000 mm/s, acceleration 3000 mm/s^2 (useActiveTCP=false optimoveEnabled=false optiMoveSpeed=0.3 optiMoveAcceleration=0.09) tcp=t0_Flange; feature=Base
          Waypoint Variable (Variable): variable=WpHome
        EvtDock := 0
Event  expression=EvtBeep
  Loop While (checkContinuously=false) expression=EvtBeep
    Set DigitalOutput pin=Do_Horn; digitalValue=1
    Set DigitalOutput pin=Do_Blue; digitalValue=1
    Wait Sleep waitTime=0.5
    Set DigitalOutput pin=Do_Horn; digitalValue=0
    Set DigitalOutput pin=Do_Blue; digitalValue=0
    Wait Sleep waitTime=5
SubProgram GripperOpen [hidden by the author, left out]
SubProgram GripperOpenQuick [hidden by the author, left out]
SubProgram GripperClose [hidden by the author, left out]
SubProgram CamAcquire (keepSynchronizedWithDisk=false)
  Folder Trig camera and process data
    Folder Init
      CamCorrectnOK := 0
      CamRetry := 0
    Wait Condition expression=SetCameraProg≟0
    Loop While (checkContinuously=false) expression=CamRetry<3
      Folder Trig
        CnxCounter := CnxAI_Counter
        Set DigitalOutput pin=CnxDO_Trig; digitalValue=1
        Timer (action=Reset) variable(name=CamTimeout)
        Timer (action=Start) variable=CamTimeout
        Wait Condition expression=CamTimeout>1 or CnxAI_Counter≠CnxCounter
        Set DigitalOutput pin=CnxDO_Trig; digitalValue=0
        Wait Sleep waitTime=0.2
        If CnxAI_Result≥100 and CnxAI_Counter≠CnxCounter
          CamRetry := 100
        Else 
          Wait Sleep waitTime=1
          CamRetry := CamRetry+1
    Folder New data validation
      If CamRetry≟100
        CamCorrectnOK := ProgExe
      Else 
        CamCorrectnOK := 0
      CamData := [(CnxAI_ResultX-30000)/10000,(CnxAI_ResultY-30000)/10000,d2r((CnxAI_ResultR-30000)/10)]
      SuppressedNode
        If CamData[1]>0.03
          Err_state := 103
      SuppressedNode
        If CamData[1]<-0.03
          Err_state := 104
      SuppressedNode
        If CamData[2]>15
          Err_state := 105
      SuppressedNode
        If CamData[2]<-15
          Err_state := 106
SubProgram GripperCloseQuick [hidden by the author, left out]
SubProgram CamCalculateCorectnPlane (keepSynchronizedWithDisk=false)
  Folder Folder
    Set NoAction tcp=t0_Flange
    Script: sync()
    P_act := get_actual_tcp_pose()
    CamCorrection := p[0,CamData[0]*-1,CamData[1],0,0,0]
    CamOffset := pose_trans(P_act,CamCorrection)
    Base_w_correctn := pose_sub(CamOffset, P_act)
